(* IEC 61131-3 sources: plc-st-coding-agent/progress/evidence/f14_p1_20261111b/jobs/codex_minimax-m27, 60 files *)

(* ---- public-easy-02.candidate_01.st ---- *)
FUNCTION_BLOCK FB_DualWordEdgeDetection
VAR_INPUT
    value : DWORD;
END_VAR

VAR_OUTPUT
    hasChanged      : BOOL;
    hasRisingEdges  : BOOL;
    risingBits      : DWORD;
    noOfRisingBits  : USINT;
    hasFallingEdges : BOOL;
    fallingBits     : DWORD;
    noOfFallingBits : USINT;
END_VAR

VAR
    prevValue : DWORD;
END_VAR

// Detect if the input value has changed
hasChanged := (value <> prevValue);

// Rising edges: current value bit is 1 AND previous value bit was 0
risingBits := value AND (NOT prevValue);
hasRisingEdges := (risingBits <> 0);

// Falling edges: current value bit is 0 AND previous value bit was 1
fallingBits := (NOT value) AND prevValue;
hasFallingEdges := (fallingBits <> 0);

// Count the number of set bits in risingBits
noOfRisingBits := 0;
IF risingBits.0 THEN noOfRisingBits := noOfRisingBits + 1; END_IF
IF risingBits.1 THEN noOfRisingBits := noOfRisingBits + 1; END_IF
IF risingBits.2 THEN noOfRisingBits := noOfRisingBits + 1; END_IF
IF risingBits.3 THEN noOfRisingBits := noOfRisingBits + 1; END_IF
IF risingBits.4 THEN noOfRisingBits := noOfRisingBits + 1; END_IF
IF risingBits.5 THEN noOfRisingBits := noOfRisingBits + 1; END_IF
IF risingBits.6 THEN noOfRisingBits := noOfRisingBits + 1; END_IF
IF risingBits.7 THEN noOfRisingBits := noOfRisingBits + 1; END_IF
IF risingBits.8 THEN noOfRisingBits := noOfRisingBits + 1; END_IF
IF risingBits.9 THEN noOfRisingBits := noOfRisingBits + 1; END_IF
IF risingBits.10 THEN noOfRisingBits := noOfRisingBits + 1; END_IF
IF risingBits.11 THEN noOfRisingBits := noOfRisingBits + 1; END_IF
IF risingBits.12 THEN noOfRisingBits := noOfRisingBits + 1; END_IF
IF risingBits.13 THEN noOfRisingBits := noOfRisingBits + 1; END_IF
IF risingBits.14 THEN noOfRisingBits := noOfRisingBits + 1; END_IF
IF risingBits.15 THEN noOfRisingBits := noOfRisingBits + 1; END_IF
IF risingBits.16 THEN noOfRisingBits := noOfRisingBits + 1; END_IF
IF risingBits.17 THEN noOfRisingBits := noOfRisingBits + 1; END_IF
IF risingBits.18 THEN noOfRisingBits := noOfRisingBits + 1; END_IF
IF risingBits.19 THEN noOfRisingBits := noOfRisingBits + 1; END_IF
IF risingBits.20 THEN noOfRisingBits := noOfRisingBits + 1; END_IF
IF risingBits.21 THEN noOfRisingBits := noOfRisingBits + 1; END_IF
IF risingBits.22 THEN noOfRisingBits := noOfRisingBits + 1; END_IF
IF risingBits.23 THEN noOfRisingBits := noOfRisingBits + 1; END_IF
IF risingBits.24 THEN noOfRisingBits := noOfRisingBits + 1; END_IF
IF risingBits.25 THEN noOfRisingBits := noOfRisingBits + 1; END_IF
IF risingBits.26 THEN noOfRisingBits := noOfRisingBits + 1; END_IF
IF risingBits.27 THEN noOfRisingBits := noOfRisingBits + 1; END_IF
IF risingBits.28 THEN noOfRisingBits := noOfRisingBits + 1; END_IF
IF risingBits.29 THEN noOfRisingBits := noOfRisingBits + 1; END_IF
IF risingBits.30 THEN noOfRisingBits := noOfRisingBits + 1; END_IF
IF risingBits.31 THEN noOfRisingBits := noOfRisingBits + 1; END_IF

// Count the number of set bits in fallingBits
noOfFallingBits := 0;
IF fallingBits.0 THEN noOfFallingBits := noOfFallingBits + 1; END_IF
IF fallingBits.1 THEN noOfFallingBits := noOfFallingBits + 1; END_IF
IF fallingBits.2 THEN noOfFallingBits := noOfFallingBits + 1; END_IF
IF fallingBits.3 THEN noOfFallingBits := noOfFallingBits + 1; END_IF
IF fallingBits.4 THEN noOfFallingBits := noOfFallingBits + 1; END_IF
IF fallingBits.5 THEN noOfFallingBits := noOfFallingBits + 1; END_IF
IF fallingBits.6 THEN noOfFallingBits := noOfFallingBits + 1; END_IF
IF fallingBits.7 THEN noOfFallingBits := noOfFallingBits + 1; END_IF
IF fallingBits.8 THEN noOfFallingBits := noOfFallingBits + 1; END_IF
IF fallingBits.9 THEN noOfFallingBits := noOfFallingBits + 1; END_IF
IF fallingBits.10 THEN noOfFallingBits := noOfFallingBits + 1; END_IF
IF fallingBits.11 THEN noOfFallingBits := noOfFallingBits + 1; END_IF
IF fallingBits.12 THEN noOfFallingBits := noOfFallingBits + 1; END_IF
IF fallingBits.13 THEN noOfFallingBits := noOfFallingBits + 1; END_IF
IF fallingBits.14 THEN noOfFallingBits := noOfFallingBits + 1; END_IF
IF fallingBits.15 THEN noOfFallingBits := noOfFallingBits + 1; END_IF
IF fallingBits.16 THEN noOfFallingBits := noOfFallingBits + 1; END_IF
IF fallingBits.17 THEN noOfFallingBits := noOfFallingBits + 1; END_IF
IF fallingBits.18 THEN noOfFallingBits := noOfFallingBits + 1; END_IF
IF fallingBits.19 THEN noOfFallingBits := noOfFallingBits + 1; END_IF
IF fallingBits.20 THEN noOfFallingBits := noOfFallingBits + 1; END_IF
IF fallingBits.21 THEN noOfFallingBits := noOfFallingBits + 1; END_IF
IF fallingBits.22 THEN noOfFallingBits := noOfFallingBits + 1; END_IF
IF fallingBits.23 THEN noOfFallingBits := noOfFallingBits + 1; END_IF
IF fallingBits.24 THEN noOfFallingBits := noOfFallingBits + 1; END_IF
IF fallingBits.25 THEN noOfFallingBits := noOfFallingBits + 1; END_IF
IF fallingBits.26 THEN noOfFallingBits := noOfFallingBits + 1; END_IF
IF fallingBits.27 THEN noOfFallingBits := noOfFallingBits + 1; END_IF
IF fallingBits.28 THEN noOfFallingBits := noOfFallingBits + 1; END_IF
IF fallingBits.29 THEN noOfFallingBits := noOfFallingBits + 1; END_IF
IF fallingBits.30 THEN noOfFallingBits := noOfFallingBits + 1; END_IF
IF fallingBits.31 THEN noOfFallingBits := noOfFallingBits + 1; END_IF

// Store current value for next cycle
prevValue := value;

END_FUNCTION_BLOCK

(* ---- public-easy-02.candidate_02.st ---- *)
FUNCTION_BLOCK FB_DualWordEdgeDetection
VAR_INPUT
    value : DWORD;
END_VAR

VAR_OUTPUT
    hasChanged      : BOOL;
    hasRisingEdges  : BOOL;
    risingBits      : DWORD;
    noOfRisingBits  : USINT;
    hasFallingEdges : BOOL;
    fallingBits     : DWORD;
    noOfFallingBits : USINT;
END_VAR

VAR
    prevValue : DWORD;
END_VAR

// Detect if the input value has changed
hasChanged := (value <> prevValue);

// Rising edges: current value bit is 1 AND previous value bit was 0
risingBits := value AND (NOT prevValue);
hasRisingEdges := (risingBits <> 0);

// Falling edges: current value bit is 0 AND previous value bit was 1
fallingBits := (NOT value) AND prevValue;
hasFallingEdges := (fallingBits <> 0);

// Count the number of set bits in risingBits using bit manipulation
noOfRisingBits := 0;
VAR tempRising : DWORD; END_VAR
tempRising := risingBits;
WHILE tempRising <> 0 DO
    noOfRisingBits := noOfRisingBits + 1;
    tempRising := tempRising AND (tempRising - 1); // Clear lowest set bit
END_WHILE

// Count the number of set bits in fallingBits using bit manipulation
noOfFallingBits := 0;
VAR tempFalling : DWORD; END_VAR
tempFalling := fallingBits;
WHILE tempFalling <> 0 DO
    noOfFallingBits := noOfFallingBits + 1;
    tempFalling := tempFalling AND (tempFalling - 1); // Clear lowest set bit
END_WHILE

// Store current value for next cycle
prevValue := value;

END_FUNCTION_BLOCK

(* ---- public-easy-03.candidate_01.st ---- *)
FUNCTION_BLOCK AlarmHandler
VAR_INPUT
    Value       : REAL;
    hiLevel     : REAL;
    loLevel     : REAL;
    hystWindow  : REAL;
END_VAR

VAR_OUTPUT
    hiAlarm     : BOOL;
    loAlarm     : BOOL;
    error       : BOOL;
    status      : WORD;
END_VAR

// Error checking
IF loLevel >= hiLevel THEN
    error := TRUE;
    status := 16#8001;
    RETURN;
END_IF

IF hystWindow >= (hiLevel - loLevel) THEN
    error := TRUE;
    status := 16#8002;
    RETURN;
END_IF

// No error
error := FALSE;
status := 16#0000;

// High alarm with hysteresis
// Trigger: Value > hiLevel
// Reset:   Value < hiLevel - hystWindow
IF Value > hiLevel THEN
    hiAlarm := TRUE;
ELSIF Value < (hiLevel - hystWindow) THEN
    hiAlarm := FALSE;
END_IF

// Low alarm with hysteresis
// Trigger: Value < loLevel
// Reset:   Value > loLevel + hystWindow
IF Value < loLevel THEN
    loAlarm := TRUE;
ELSIF Value > (loLevel + hystWindow) THEN
    loAlarm := FALSE;
END_IF

END_FUNCTION_BLOCK

(* ---- public-easy-03.candidate_02.st ---- *)
FUNCTION_BLOCK AlarmHandler
VAR_INPUT
    Value       : REAL;
    hiLevel     : REAL;
    loLevel     : REAL;
    hystWindow  : REAL;
END_VAR

VAR_OUTPUT
    hiAlarm     : BOOL;
    loAlarm     : BOOL;
    error       : BOOL;
    status      : WORD;
END_VAR

// Error checking
IF loLevel >= hiLevel THEN
    error := TRUE;
    status := 16#8001;
    RETURN;
END_IF

IF hystWindow >= (hiLevel - loLevel) THEN
    error := TRUE;
    status := 16#8002;
    RETURN;
END_IF

// No error - reset all outputs to defined state
error := FALSE;
status := 16#0000;
hiAlarm := FALSE;
loAlarm := FALSE;

// High alarm with hysteresis
// Trigger: Value > hiLevel
// Reset:   Value < hiLevel - hystWindow
IF Value > hiLevel THEN
    hiAlarm := TRUE;
END_IF

// Low alarm with hysteresis
// Trigger: Value < loLevel
// Reset:   Value > loLevel + hystWindow
IF Value < loLevel THEN
    loAlarm := TRUE;
END_IF

END_FUNCTION_BLOCK

(* ---- public-easy-05.candidate_01.st ---- *)
FUNCTION_BLOCK WeldGapAlarm
VAR_INPUT
    Gap_Exceeded    : BOOL;      // Scanner indication that the gap exceeds 1.5 mm
    Weld_E_Stop_NC  : BOOL;      // TRUE = inactive, FALSE = active (emergency stop)
    DebounceTime    : TIME;      // Gap-signal debounce duration during normal monitoring
END_VAR

VAR_OUTPUT
    Operator_Alert         : BOOL;  // Audible and visual alarm command
    Weld_Soft_Start_Active : BOOL;  // Monitoring-inhibition status during 5-second power-up initialization
END_VAR

VAR
    InitTimer    : TON;          // 5-second initialization inhibition timer
    DebounceTmr  : TON;          // Gap signal debounce timer during normal monitoring
    bInitDone    : BOOL;         // Power-up initialization completion flag
END_VAR

    // E-Stop takes highest priority over initialization and normal monitoring
    IF NOT Weld_E_Stop_NC THEN
        Operator_Alert         := FALSE;
        Weld_Soft_Start_Active := FALSE;
        DebounceTmr(IN := FALSE);
        InitTimer(IN := FALSE);
        bInitDone := FALSE;
        RETURN;
    END_IF

    // 5-second initialization inhibition period
    IF NOT bInitDone THEN
        Weld_Soft_Start_Active := TRUE;
        Operator_Alert         := FALSE;
        InitTimer(IN := TRUE, PT := T#5S);

        IF InitTimer.Q THEN
            bInitDone := TRUE;
            InitTimer(IN := FALSE);
        END_IF;

        // During initialization, debounce time does NOT accumulate
        RETURN;
    END_IF;

    // Normal gap monitoring after initialization
    Weld_Soft_Start_Active := FALSE;

    // Debounce logic: alarm only after Gap_Exceeded remains TRUE for DebounceTime
    IF Gap_Exceeded THEN
        DebounceTmr(IN := TRUE, PT := DebounceTime);
        Operator_Alert := DebounceTmr.Q;
    ELSE
        DebounceTmr(IN := FALSE);
        Operator_Alert := FALSE;
    END_IF;

END_FUNCTION_BLOCK

(* ---- public-easy-05.candidate_02.st ---- *)
FUNCTION_BLOCK WeldGapAlarm
VAR_INPUT
    Gap_Exceeded    : BOOL;      // Scanner indication that the gap exceeds 1.5 mm
    Weld_E_Stop_NC  : BOOL;      // TRUE = inactive, FALSE = active (emergency stop)
    DebounceTime    : TIME;      // Gap-signal debounce duration during normal monitoring
END_VAR

VAR_OUTPUT
    Operator_Alert         : BOOL;  // Audible and visual alarm command
    Weld_Soft_Start_Active : BOOL;  // Monitoring-inhibition status during 5-second power-up initialization
END_VAR

VAR
    InitTimer    : TON;          // 5-second initialization inhibition timer
    DebounceTmr  : TON;          // Gap signal debounce timer during normal monitoring
    bInitDone    : BOOL;         // Power-up initialization completion flag
END_VAR

    // E-Stop takes highest priority over initialization and normal monitoring
    IF NOT Weld_E_Stop_NC THEN
        Operator_Alert         := FALSE;
        Weld_Soft_Start_Active := FALSE;
        DebounceTmr(IN := FALSE, R := TRUE);
        InitTimer(IN := FALSE, R := TRUE);
        bInitDone := FALSE;
        RETURN;
    END_IF

    // 5-second initialization inhibition period
    IF NOT bInitDone THEN
        Weld_Soft_Start_Active := TRUE;
        Operator_Alert         := FALSE;
        InitTimer(IN := TRUE, PT := T#5S);

        IF InitTimer.Q THEN
            bInitDone := TRUE;
            InitTimer(IN := FALSE);
        END_IF;

        // During initialization, debounce time does NOT accumulate
        RETURN;
    END_IF;

    // Normal gap monitoring after initialization
    Weld_Soft_Start_Active := FALSE;

    // Debounce logic: alarm only after Gap_Exceeded remains TRUE for DebounceTime
    IF Gap_Exceeded THEN
        DebounceTmr(IN := TRUE, PT := DebounceTime);
        Operator_Alert := DebounceTmr.Q;
    ELSE
        DebounceTmr(IN := FALSE, PT := DebounceTime);  // Reset timer to clear accumulated time
        Operator_Alert := FALSE;
    END_IF;

END_FUNCTION_BLOCK

(* ---- public-easy-06.candidate_02.st ---- *)
FUNCTION_BLOCK AerationBlower
VAR_INPUT
    do_low               : BOOL;
    aeration_e_stop_nc   : BOOL;
END_VAR

VAR_OUTPUT
    blower_run                   : BOOL;
    aeration_blower_cycle_count  : UINT;
END_VAR

VAR
    start_timer        : TON;
    blower_was_running : BOOL;
END_VAR

// Start delay: timer runs while both conditions are met
start_timer(
    IN := do_low AND aeration_e_stop_nc,
    PT := T#5S
);

// Blower runs only when timer elapsed AND conditions remain satisfied
blower_run := start_timer.Q AND do_low AND aeration_e_stop_nc;

// Count FALSE-to-TRUE transitions of blower_run (rising edge)
IF blower_run AND NOT blower_was_running THEN
    aeration_blower_cycle_count := aeration_blower_cycle_count + 1;
END_IF;

// Update edge-detection state for next scan
blower_was_running := blower_run;

END_FUNCTION_BLOCK

(* ---- public-hard-01.candidate_02.st ---- *)
// Material Proportioning Process Control - ST Implementation
FUNCTION_BLOCK MaterialProportioning
VAR_INPUT
    estop            : BOOL;   // Emergency Stop Signal (FALSE = triggered)
    opeMode          : BOOL;   // Operation Mode (FALSE = Manual, TRUE = Auto)
    valveAStart      : BOOL;   // Valve A Start Button
    valveBStart      : BOOL;   // Valve B Start Button
    valveCStart      : BOOL;   // Valve C Start Button
    valveDStart      : BOOL;   // Valve D Start Button
    mixMotorStart    : BOOL;   // Mixing Motor Start Button
    autoStart        : BOOL;   // Automatic Start Button
    processMode      : BOOL;   // Process Mode (FALSE = Basic, TRUE = Extended)
    levelSensor      : INT;    // Liquid Level Sensor (unit: cm)
    mixMotorComplete : BOOL;   // Mixing Complete Signal
END_VAR

VAR_OUTPUT
    valveARun  : BOOL;   // Valve A Run Command
    valveBRun  : BOOL;   // Valve B Run Command
    valveCRun  : BOOL;   // Valve C Run Command
    valveDRun  : BOOL;   // Valve D Run Command
    mixMotorRun: BOOL;   // Mixing Motor Run Command
END_VAR

VAR
    prevValveAStart   : BOOL;   // Previous state for edge detection
    prevValveBStart   : BOOL;
    prevValveCStart   : BOOL;
    prevValveDStart   : BOOL;
    prevMixMotorStart : BOOL;
    prevAutoStart     : BOOL;
    autoState : INT;     // 0=IDLE, 1=FILL_A, 2=FILL_B, 3=MIX_BASIC,
                         // 4=FILL_C, 5=MIX_EXT, 6=DRAIN
END_VAR

VAR CONSTANT
    STATE_IDLE      : INT := 0;
    STATE_FILL_A    : INT := 1;
    STATE_FILL_B    : INT := 2;
    STATE_MIX_BASIC : INT := 3;
    STATE_FILL_C    : INT := 4;
    STATE_MIX_EXT   : INT := 5;
    STATE_DRAIN     : INT := 6;
END_VAR

// ============================================================================
// Main Control Logic
// ============================================================================

// ---------------------------------------------------------------------------
// Emergency Stop Logic
// When estop=FALSE, all equipment stops immediately
// ---------------------------------------------------------------------------
IF NOT estop THEN
    valveARun  := FALSE;
    valveBRun  := FALSE;
    valveCRun  := FALSE;
    valveDRun  := FALSE;
    mixMotorRun:= FALSE;
    autoState  := STATE_IDLE;

    prevValveAStart   := FALSE;
    prevValveBStart   := FALSE;
    prevValveCStart   := FALSE;
    prevValveDStart   := FALSE;
    prevMixMotorStart := FALSE;
    prevAutoStart     := FALSE;
    RETURN;
END_IF

// ---------------------------------------------------------------------------
// Mode Selection: Manual vs Automatic
// ---------------------------------------------------------------------------
IF NOT opeMode THEN
    // MANUAL OPERATION MODE
    // Toggle each device on rising edge of corresponding button

    IF valveAStart AND NOT prevValveAStart THEN
        valveARun := NOT valveARun;
    END_IF;
    prevValveAStart := valveAStart;

    IF valveBStart AND NOT prevValveBStart THEN
        valveBRun := NOT valveBRun;
    END_IF;
    prevValveBStart := valveBStart;

    IF valveCStart AND NOT prevValveCStart THEN
        valveCRun := NOT valveCRun;
    END_IF;
    prevValveCStart := valveCStart;

    IF valveDStart AND NOT prevValveDStart THEN
        valveDRun := NOT valveDRun;
    END_IF;
    prevValveDStart := valveDStart;

    IF mixMotorStart AND NOT prevMixMotorStart THEN
        mixMotorRun := NOT mixMotorRun;
    END_IF;
    prevMixMotorStart := mixMotorStart;

ELSE
    // AUTOMATIC OPERATION MODE

    valveARun  := FALSE;
    valveBRun  := FALSE;
    valveCRun  := FALSE;
    valveDRun  := FALSE;
    mixMotorRun:= FALSE;

    IF autoStart AND NOT prevAutoStart THEN
        IF autoState = STATE_IDLE THEN
            autoState := STATE_FILL_A;
        END_IF;
    END_IF;
    prevAutoStart := autoStart;

    CASE autoState OF

        STATE_IDLE:
            valveARun  := FALSE;
            valveBRun  := FALSE;
            valveCRun  := FALSE;
            valveDRun  := FALSE;
            mixMotorRun:= FALSE;

        STATE_FILL_A:
            valveARun := TRUE;
            IF levelSensor >= 50 THEN
                valveARun := FALSE;
                autoState := STATE_FILL_B;
            END_IF;

        STATE_FILL_B:
            valveBRun := TRUE;
            IF levelSensor >= 80 THEN
                valveBRun := FALSE;
                IF NOT processMode THEN
                    autoState := STATE_MIX_BASIC;
                ELSE
                    autoState := STATE_FILL_C;
                END_IF;
            END_IF;

        STATE_MIX_BASIC:
            mixMotorRun := TRUE;
            IF mixMotorComplete THEN
                mixMotorRun := FALSE;
                autoState := STATE_DRAIN;
            END_IF;

        STATE_FILL_C:
            valveCRun := TRUE;
            IF levelSensor >= 100 THEN
                valveCRun := FALSE;
                autoState := STATE_MIX_EXT;
            END_IF;

        STATE_MIX_EXT:
            mixMotorRun := TRUE;
            IF mixMotorComplete THEN
                mixMotorRun := FALSE;
                autoState := STATE_DRAIN;
            END_IF;

        STATE_DRAIN:
            valveDRun := TRUE;
            IF levelSensor < 10 THEN
                valveDRun := FALSE;
                autoState := STATE_IDLE;
            END_IF;

    END_CASE;

END_IF;

END_FUNCTION_BLOCK

PROGRAM PLC_PRG
VAR
    inst : MaterialProportioning;
END_VAR

inst(
    estop            := estop,
    opeMode          := opeMode,
    valveAStart      := valveAStart,
    valveBStart      := valveBStart,
    valveCStart      := valveCStart,
    valveDStart      := valveDStart,
    mixMotorStart    := mixMotorStart,
    autoStart        := autoStart,
    processMode      := processMode,
    levelSensor      := levelSensor,
    mixMotorComplete := mixMotorComplete,
    valveARun        => valveARun,
    valveBRun        => valveBRun,
    valveCRun        => valveCRun,
    valveDRun        => valveDRun,
    mixMotorRun      => mixMotorRun
);
END_PROGRAM

(* ---- public-hard-04.candidate_02.st ---- *)
FUNCTION_BLOCK FB_FIFO
VAR_INPUT
    enqueue : BOOL;
    dequeue : BOOL;
    reset   : BOOL;
END_VAR

VAR_OUTPUT
    elementCount : DINT;
    status       : WORD;
END_VAR

VAR_IN_OUT
    item   : VARIANT;
    buffer : VARIANT;
END_VAR

VAR
    _head         : DINT := 0;
    _tail         : DINT := 0;
    _elementCount : DINT := 0;
    _capacity     : DINT;
    _elementSize  : DINT;
    _prevEnqueue  : BOOL := FALSE;
    _prevDequeue  : BOOL := FALSE;
    _initialized  : BOOL := FALSE;
END_VAR

// Initialization
IF NOT _initialized THEN
    VAR
        bufType : REF_TO ANY;
        capacity : DINT;
    END_VAR

    bufType REF= buffer;

    IF __ISVALIDREF(bufType) THEN
        capacity := bufType.GetUpperBound(1) + 1;
        _capacity := capacity;
        _elementSize := bufType.GetSize() / _capacity;
        _initialized := TRUE;
    END_IF;

    elementCount := 0;
    status := 16#0000;
    RETURN;
END_IF;

// Reset handling (highest priority)
IF reset THEN
    _head := 0;
    _tail := 0;
    _elementCount := 0;
    elementCount := 0;
    status := 16#0000;
    _prevEnqueue := FALSE;
    _prevDequeue := FALSE;
    RETURN;
END_IF;

// Rising edge detection
VAR
    enqueueRising : BOOL;
    dequeueRising : BOOL;
END_VAR

enqueueRising := enqueue AND NOT _prevEnqueue;
dequeueRising := dequeue AND NOT _prevDequeue;

_prevEnqueue := enqueue;
_prevDequeue := dequeue;

// Dequeue request (rising edge, queue not empty)
IF dequeueRising AND _elementCount > 0 THEN
    VAR
        pSrc     : POINTER TO BYTE;
        pDest    : POINTER TO BYTE;
        srcAdr   : LWORD;
        destAdr  : LWORD;
        zeroBuf  : ARRAY[0..255] OF BYTE;
    END_VAR

    srcAdr := __GET_VAR_DATA_REF(buffer).ADR + (_head * _elementSize);
    destAdr := __GET_VAR_DATA_REF(item).ADR;

    MemMove(TO_PTR(srcAdr), TO_PTR(destAdr), _elementSize);

    MemSet(zeroBuf, 0, SIZEOF(zeroBuf));
    MemMove(zeroBuf, TO_PTR(srcAdr), _elementSize);

    _head := (_head + 1) MOD _capacity;
    _elementCount := _elementCount - 1;
    elementCount := _elementCount;
    status := 16#0000;

// Enqueue request (rising edge, queue not full)
ELSIF enqueueRising AND _elementCount < _capacity THEN
    VAR
        pDest   : POINTER TO BYTE;
        pSrc    : POINTER TO BYTE;
        destAdr : LWORD;
        srcAdr  : LWORD;
    END_VAR

    destAdr := __GET_VAR_DATA_REF(buffer).ADR + (_tail * _elementSize);
    srcAdr := __GET_VAR_DATA_REF(item).ADR;

    MemMove(TO_PTR(srcAdr), TO_PTR(destAdr), _elementSize);

    _tail := (_tail + 1) MOD _capacity;
    _elementCount := _elementCount + 1;
    elementCount := _elementCount;
    status := 16#0000;

// Dequeue rejected: empty queue
ELSIF dequeueRising AND _elementCount = 0 THEN
    status := 16#8001;

// Enqueue rejected: full queue
ELSIF enqueueRising AND _elementCount >= _capacity THEN
    status := 16#8002;

// Idle (no rising edge or other condition)
ELSE
    status := 16#0000;
END_IF;
END_FUNCTION_BLOCK

(* ---- public-medium-01.candidate_02.st ---- *)
FUNCTION_BLOCK FB_MultiPumpControl
VAR_INPUT
    mode    : BOOL;  // FALSE: Manual mode, TRUE: Automatic mode
    start   : BOOL;  // Start button
    stop    : BOOL;  // Stop button
END_VAR

VAR_IN_OUT
    pumpGroup   : ARRAY[1..5] OF ST_Pump;
END_VAR

VAR
    startOld    : BOOL := FALSE;
    stopOld     : BOOL := FALSE;
    startEdge   : BOOL;
    stopEdge    : BOOL;
    i           : INT;
    runCount    : INT;
    tempPump    : ST_Pump;
    sorted      : BOOL := FALSE;
    priorities  : ARRAY[1..5] OF INT;
END_VAR

// Detect rising edges
startEdge := start AND NOT startOld;
stopEdge  := stop  AND NOT stopOld;
startOld  := start;
stopOld   := stop;

// Stop all pumps when stop is pressed
IF stopEdge THEN
    FOR i := 1 TO 5 DO
        pumpGroup[i].RunComd := FALSE;
    END_FOR
    sorted := FALSE;
    RETURN;
END_IF

// Start pumps when start is pressed
IF startEdge THEN
    IF mode = FALSE THEN
        // Manual mode: start pumps based on selection
        FOR i := 1 TO 5 DO
            IF pumpGroup[i].selection THEN
                pumpGroup[i].RunComd := TRUE;
            END_IF
        END_FOR
    ELSE
        // Automatic mode: select top 3 by priority (bubble sort)
        // Store priorities
        FOR i := 1 TO 5 DO
            priorities[i] := pumpGroup[i].priority;
        END_FOR

        // Bubble sort priorities and rearrange pumpGroup accordingly
        FOR i := 1 TO 5 DO
            tempPump := pumpGroup[i];
        END_FOR

        // Sort by priority descending
        FOR i := 1 TO 4 DO
            IF priorities[i] < priorities[i+1] THEN
                // Swap priorities
                tempPump := pumpGroup[i];
                pumpGroup[i] := pumpGroup[i+1];
                pumpGroup[i+1] := tempPump;

                // Update priority array
                priorities[i] := pumpGroup[i].priority;
                priorities[i+1] := pumpGroup[i+1].priority;
            END_IF
        END_FOR

        // Select top 3 pumps
        runCount := 0;
        FOR i := 1 TO 5 DO
            IF runCount < 3 THEN
                pumpGroup[i].RunComd := TRUE;
                runCount := runCount + 1;
            ELSE
                pumpGroup[i].RunComd := FALSE;
            END_IF
        END_FOR

        sorted := TRUE;
    END_IF
END_IF
END_FUNCTION_BLOCK

(* ---- public-medium-02.candidate_01.st ---- *)
FUNCTION_BLOCK FB_AnalogBatchProcess
VAR_INPUT
    count : DINT;
END_VAR

VAR_IN_OUT
    analogValues : ARRAY[*] OF INT;
    channels     : ARRAY[*] OF ST_AnalogChannel;
END_VAR

VAR
    i           : DINT;
    idx         : DINT;
    rawValue    : INT;
    channel     : REF_TO ST_AnalogChannel;
END_VAR

// Process each channel by ordinal position
FOR i := 0 TO count - 1 DO
    idx := LOWER_BOUND(channels, 1) + i;
    channel := REF(channels[idx]);

    // Skip disabled channels
    IF NOT channel.enable THEN
        CONTINUE;
    END_IF

    // Default success status
    channel.retVal := 16#0000;

    // Validate hiLIM > loLIM
    IF channel.hiLIM <= channel.loLIM THEN
        channel.retVal := 16#8002;
        CONTINUE;
    END_IF

    // Get raw analog value (read-only)
    rawValue := analogValues[LOWER_BOUND(analogValues, 1) + i];

    // Perform conversion based on measuringMode
    CASE channel.measuringMode OF
        0: // Non-temperature linear scaling
            IF channel.bipolar THEN
                // Bipolar: map -27648..27648 to loLIM..hiLIM
                channel.outputValue := (INT_TO_REAL(rawValue) + 27648.0) / 55296.0 * (channel.hiLIM - channel.loLIM) + channel.loLIM;
            ELSE
                // Unipolar: map 0..27648 to loLIM..hiLIM
                channel.outputValue := INT_TO_REAL(rawValue) / 27648.0 * (channel.hiLIM - channel.loLIM) + channel.loLIM;
            END_IF;

        1: // Standard temperature: outputValue = raw / 10
            channel.outputValue := INT_TO_REAL(rawValue) / 10.0;

        2: // Climatic temperature: outputValue = raw / 100
            channel.outputValue := INT_TO_REAL(rawValue) / 100.0;

    ELSE
        // Invalid measuringMode
        channel.retVal := 16#8001;
    END_CASE;
END_FOR;

END_FUNCTION_BLOCK

(* ---- public-medium-02.candidate_02.st ---- *)
FUNCTION_BLOCK FB_AnalogBatchProcess
VAR_INPUT
    count : DINT;
END_VAR

VAR_IN_OUT
    analogValues : ARRAY[*] OF INT;
    channels     : ARRAY[*] OF ST_AnalogChannel;
END_VAR

VAR
    i           : DINT;
    idx         : DINT;
    rawValue    : INT;
    validInput  : BOOL;
END_VAR

i := 0;
WHILE i < count DO
    idx := LOWER_BOUND(channels, 1) + i;

    // Check if channel is enabled
    IF channels[idx].enable THEN
        // Default success status
        channels[idx].retVal := 16#0000;

        // Validate hiLIM > loLIM
        IF channels[idx].hiLIM > channels[idx].loLIM THEN
            // Get raw analog value
            rawValue := analogValues[LOWER_BOUND(analogValues, 1) + i];

            // Perform conversion based on measuringMode
            CASE channels[idx].measuringMode OF
                0: // Non-temperature linear scaling
                    IF channels[idx].bipolar THEN
                        // Bipolar: map -27648..27648 to loLIM..hiLIM
                        channels[idx].outputValue := (INT_TO_REAL(rawValue) + 27648.0) / 55296.0 * (channels[idx].hiLIM - channels[idx].loLIM) + channels[idx].loLIM;
                    ELSE
                        // Unipolar: map 0..27648 to loLIM..hiLIM
                        channels[idx].outputValue := INT_TO_REAL(rawValue) / 27648.0 * (channels[idx].hiLIM - channels[idx].loLIM) + channels[idx].loLIM;
                    END_IF;

                1: // Standard temperature: outputValue = raw / 10
                    channels[idx].outputValue := INT_TO_REAL(rawValue) / 10.0;

                2: // Climatic temperature: outputValue = raw / 100
                    channels[idx].outputValue := INT_TO_REAL(rawValue) / 100.0;

            ELSE
                // Invalid measuringMode
                channels[idx].retVal := 16#8001;
            END_CASE;
        ELSE
            // hiLIM <= loLIM error
            channels[idx].retVal := 16#8002;
        END_IF;
    END_IF;

    i := i + 1;
END_WHILE;

END_FUNCTION_BLOCK

(* ---- public-medium-04.candidate_01.st ---- *)
FUNCTION_BLOCK FB_TemperatureControl
VAR_INPUT
    TemperatureSensorInput : REAL;
    SetTemperature         : REAL;
END_VAR

VAR_OUTPUT
    CurrentTemperature : REAL;
    SetTempDisplay     : REAL;
    HeaterStatus       : BOOL;
    OverheatProtection : BOOL;
    HeaterOutput       : BOOL;
END_VAR

VAR
    // Internal variables
    rCurrentTemperature  : REAL := 0.0;
    rSetTemperature      : REAL := 0.0;
    bHeaterOn            : BOOL := FALSE;
    bOverheatProtection  : BOOL := FALSE;
    bSensorFault         : BOOL := FALSE;

    // Timer for heater on-time monitoring
    HeaterOnTimer        : TON;
    // Timer for overheat protection cooldown
    OverheatCooldownTimer: TON;

    // Constants
    MAX_HEATER_ON_TIME   : TIME := T#5S;
    OVERHEAT_COOLDOWN    : TIME := T#3S;
    MIN_SENSOR_VALUE     : REAL := 0.0;
    MAX_SENSOR_VALUE     : REAL := 100.0;
END_VAR

//============================================================================
// Temperature Logic Control - Main Program
//============================================================================

// Update internal temperature values from inputs
rCurrentTemperature := TemperatureSensorInput;
rSetTemperature     := SetTemperature;

// Update output displays
CurrentTemperature := rCurrentTemperature;
SetTempDisplay     := rSetTemperature;
HeaterStatus       := bHeaterOn;
OverheatProtection := bOverheatProtection;

//============================================================================
// Sensor Fault Detection
// If temperature is outside valid range (0-100), trigger sensor fault
//============================================================================
bSensorFault := (rCurrentTemperature < MIN_SENSOR_VALUE) OR
                (rCurrentTemperature > MAX_SENSOR_VALUE);

IF bSensorFault THEN
    // Sensor fault: turn off heater immediately
    bHeaterOn          := FALSE;
    HeaterOutput       := FALSE;
    bOverheatProtection := TRUE;

    // Reset heater on timer when heater is off
    HeaterOnTimer(IN := FALSE);

    // Return early - no temperature control during sensor fault
    RETURN;
END_IF;

//============================================================================
// Overheat Protection Check
// If protection is active, must wait for cooldown period before reset
//============================================================================
IF bOverheatProtection THEN
    // Start or continue cooldown timer
    OverheatCooldownTimer(IN := TRUE, PT := OVERHEAT_COOLDOWN);

    // Check if cooldown period has elapsed
    IF OverheatCooldownTimer.Q THEN
        // Cooldown complete - reset overheat protection
        bOverheatProtection        := FALSE;
        OverheatCooldownTimer(IN := FALSE);
    END_IF;

    // Keep heater off during overheat protection
    bHeaterOn := FALSE;
    HeaterOutput := FALSE;

    // Return early - no temperature control during overheat protection
    RETURN;
ELSE
    // Reset cooldown timer when protection is not active
    OverheatCooldownTimer(IN := FALSE);
END_IF;

//============================================================================
// Temperature Control Logic
// Compare actual temperature with set temperature
//============================================================================
IF rCurrentTemperature < rSetTemperature THEN
    // Temperature below setpoint - turn ON heater
    bHeaterOn := TRUE;
ELSIF rCurrentTemperature >= rSetTemperature THEN
    // Temperature at or above setpoint - turn OFF heater
    bHeaterOn := FALSE;
END_IF;

//============================================================================
// Heater Output Control
//============================================================================
HeaterOutput := bHeaterOn;

//============================================================================
// Heater On-Time Monitoring for Overheat Protection
// If heater runs continuously for more than 5 seconds, trigger protection
//============================================================================
IF bHeaterOn THEN
    // Start or continue the heater on-time timer
    HeaterOnTimer(IN := TRUE, PT := MAX_HEATER_ON_TIME);

    // Check if timer has elapsed (heater on for too long)
    IF HeaterOnTimer.Q THEN
        // Overheat protection triggered
        bHeaterOn           := FALSE;
        bOverheatProtection := TRUE;
        HeaterOutput        := FALSE;

        // Reset heater on timer
        HeaterOnTimer(IN := FALSE);
    END_IF;
ELSE
    // Heater is off - reset the timer
    HeaterOnTimer(IN := FALSE);
END_IF;

END_FUNCTION_BLOCK

(* ---- public-medium-04.candidate_02.st ---- *)
FUNCTION_BLOCK FB_TemperatureControl
VAR_INPUT
    TemperatureSensorInput : REAL;
    SetTemperature         : REAL;
END_VAR

VAR_OUTPUT
    CurrentTemperature : REAL;
    SetTempDisplay     : REAL;
    HeaterStatus       : BOOL;
    OverheatProtection : BOOL;
    HeaterOutput       : BOOL;
END_VAR

VAR
    bHeaterOn            : BOOL := FALSE;
    bOverheatProtection  : BOOL := FALSE;

    HeaterOnTimer        : TON;
    OverheatCooldownTimer: TON;

    MAX_HEATER_ON_TIME   : TIME := T#5S;
    OVERHEAT_COOLDOWN    : TIME := T#3S;
END_VAR

//============================================================================
// Main Control Logic
//============================================================================

// Sensor Fault Detection (0-100 valid range)
IF (TemperatureSensorInput < 0.0) OR (TemperatureSensorInput > 100.0) THEN
    // Sensor fault: disable heater and activate protection
    bHeaterOn := FALSE;
    bOverheatProtection := TRUE;
    HeaterOnTimer(IN := FALSE);
END_IF

// Overheat Protection Logic
IF bOverheatProtection THEN
    OverheatCooldownTimer(IN := TRUE, PT := OVERHEAT_COOLDOWN);

    IF OverheatCooldownTimer.Q THEN
        bOverheatProtection := FALSE;
        OverheatCooldownTimer(IN := FALSE);
    END_IF;

    bHeaterOn := FALSE;
ELSE
    OverheatCooldownTimer(IN := FALSE);

    // Temperature Control (only when no protection active)
    IF TemperatureSensorInput < SetTemperature THEN
        bHeaterOn := TRUE;
    ELSE
        bHeaterOn := FALSE;
    END_IF;
END_IF;

// Heater On-Time Monitoring
IF bHeaterOn THEN
    HeaterOnTimer(IN := TRUE, PT := MAX_HEATER_ON_TIME);

    IF HeaterOnTimer.Q THEN
        bHeaterOn := FALSE;
        bOverheatProtection := TRUE;
        HeaterOnTimer(IN := FALSE);
    END_IF;
ELSE
    HeaterOnTimer(IN := FALSE);
END_IF;

//============================================================================
// Update All Outputs (at the end, after all logic)
//============================================================================
CurrentTemperature := TemperatureSensorInput;
SetTempDisplay     := SetTemperature;
HeaterStatus       := bHeaterOn;
OverheatProtection := bOverheatProtection;
HeaterOutput       := bHeaterOn;

END_FUNCTION_BLOCK

(* ---- public-medium-06.candidate_02.st ---- *)
FUNCTION_BLOCK SlabThicknessMonitor
VAR_INPUT
    THICKNESS_FAULT        : BOOL;
    THICKNESS_SIGNAL_VALID : BOOL;
    cutting_run            : BOOL;
    faulttimestamp         : DINT;
    cycletime              : TIME;
END_VAR

VAR_OUTPUT
    THICKNESS_ALARM           : BOOL;
    slab_fault_counter        : UINT;
    slab_runtime_accumulator  : LTIME;
    slab_fault_history        : ARRAY[0..4] OF DINT;
END_VAR

VAR
    AlarmHoldTimer   : TON;
    FaultWasActive   : BOOL;
    PowerUpComplete  : BOOL;
    i                : INT;
END_VAR

IF NOT PowerUpComplete THEN
    THICKNESS_ALARM           := FALSE;
    slab_fault_counter        := 0;
    slab_runtime_accumulator  := LTIME#0s;

    FOR i := 0 TO 4 DO
        slab_fault_history[i] := 0;
    END_FOR

    FaultWasActive  := FALSE;
    PowerUpComplete := TRUE;
END_IF

IF NOT THICKNESS_SIGNAL_VALID THEN
    THICKNESS_ALARM := FALSE;
    AlarmHoldTimer(IN := FALSE);
    FaultWasActive  := FALSE;
ELSE
    AlarmHoldTimer(IN := THICKNESS_FAULT, PT := T#500ms);
    THICKNESS_ALARM := THICKNESS_FAULT OR AlarmHoldTimer.Q;

    IF THICKNESS_FAULT AND NOT FaultWasActive THEN
        slab_fault_counter        := slab_fault_counter + 1;
        slab_fault_history[4]     := slab_fault_history[3];
        slab_fault_history[3]     := slab_fault_history[2];
        slab_fault_history[2]     := slab_fault_history[1];
        slab_fault_history[1]     := slab_fault_history[0];
        slab_fault_history[0]     := faulttimestamp;
    END_IF;

    FaultWasActive := THICKNESS_FAULT;

    IF cutting_run AND NOT THICKNESS_FAULT THEN
        slab_runtime_accumulator := slab_runtime_accumulator + cycletime;
    END_IF
END_IF

END_FUNCTION_BLOCK

(* ---- public-medium-07.candidate_02.st ---- *)
FUNCTION_BLOCK HVAC_Control
VAR_INPUT
    OCCUPANCY_DETECTED    : BOOL;
    ENERGY_SAVING_MODE    : BOOL;
    HVAC_MODE_SELECTOR    : INT;
END_VAR

VAR_OUTPUT
    SUPPLY_FAN_RUN        : BOOL := FALSE;
    TEMP_SETPOINT_ADJUST  : INT := 0;
END_VAR

VAR
    occupancy_delay_timer : TON;
END_VAR

// Fan control with 30-second delay
IF OCCUPANCY_DETECTED AND (HVAC_MODE_SELECTOR <> 3) THEN
    occupancy_delay_timer(IN := TRUE, PT := T#30S);
    IF occupancy_delay_timer.Q THEN
        SUPPLY_FAN_RUN := TRUE;
    ELSE
        SUPPLY_FAN_RUN := FALSE;
    END_IF;
ELSE
    occupancy_delay_timer(IN := FALSE);
    SUPPLY_FAN_RUN := FALSE;
END_IF;

// Temperature setpoint adjustment per mode
CASE HVAC_MODE_SELECTOR OF
    0: // Auto
        IF OCCUPANCY_DETECTED THEN
            TEMP_SETPOINT_ADJUST := 0;
        ELSE
            TEMP_SETPOINT_ADJUST := BOOL_TO_INT(ENERGY_SAVING_MODE) + 2;
        END_IF;
    1: // Comfort
        IF OCCUPANCY_DETECTED THEN
            TEMP_SETPOINT_ADJUST := 0;
        ELSE
            TEMP_SETPOINT_ADJUST := 1;
        END_IF;
    2: // Economy
        IF OCCUPANCY_DETECTED THEN
            TEMP_SETPOINT_ADJUST := 0;
        ELSE
            TEMP_SETPOINT_ADJUST := 4;
        END_IF;
    3: // Night
        TEMP_SETPOINT_ADJUST := 4;
    ELSE
        TEMP_SETPOINT_ADJUST := 0;
END_CASE;

// Clamp to ±4°C
IF TEMP_SETPOINT_ADJUST > 4 THEN
    TEMP_SETPOINT_ADJUST := 4;
ELSIF TEMP_SETPOINT_ADJUST < -4 THEN
    TEMP_SETPOINT_ADJUST := -4;
END_IF;

END_FUNCTION_BLOCK

(* ---- public-medium-08.candidate_01.st ---- *)
FUNCTION_BLOCK FB_IPv4Parse
    VAR_INPUT
        ipText : STRING(254);
    END_VAR
    VAR_OUTPUT
        ipValue : UDINT;
    END_VAR
    VAR
        pos : INT;
        segmentStart : INT;
        segmentLen : INT;
        segmentCount : INT;
        value : INT;
        ch : CHAR;
        textLen : INT;
    END_VAR

    ipValue := 0;
    textLen := LEN(ipText);
    pos := 1;
    segmentCount := 0;

    // Skip leading whitespace
    WHILE (pos <= textLen) AND (MID(ipText, 1, pos) = ' ') DO
        pos := pos + 1;
    END_WHILE;

    // Parse up to 4 segments
    WHILE (segmentCount < 4) AND (pos <= textLen) DO
        segmentStart := pos;
        segmentLen := 0;

        // Collect digits for current segment
        WHILE (pos <= textLen) DO
            ch := MID(ipText, 1, pos);
            IF ch = '.' THEN
                EXIT;
            END_IF;
            IF (ch < '0') OR (ch > '9') THEN
                ipValue := 0;
                RETURN;
            END_IF;
            segmentLen := segmentLen + 1;
            pos := pos + 1;
        END_WHILE;

        // Check segment length (1-3 digits for valid 0-255)
        IF segmentLen < 1 OR segmentLen > 3 THEN
            ipValue := 0;
            RETURN;
        END_IF;

        // Parse segment value
        value := 0;
        FOR pos := segmentStart TO segmentStart + segmentLen - 1 DO
            ch := MID(ipText, 1, pos);
            value := value * 10 + (ch - '0');
        END_FOR;

        // Validate segment range
        IF value > 255 THEN
            ipValue := 0;
            RETURN;
        END_IF;

        // Accumulate result in network byte order
        ipValue := (ipValue << 8) OR TO_UDINT(value);
        segmentCount := segmentCount + 1;

        // Skip the dot separator if present
        IF (pos <= textLen) AND (MID(ipText, 1, pos) = '.') THEN
            pos := pos + 1;
        END_IF;
    END_WHILE;

    // Validate we have exactly 4 segments
    IF segmentCount <> 4 THEN
        ipValue := 0;
        RETURN;
    END_IF;

    // Skip trailing whitespace
    WHILE (pos <= textLen) AND (MID(ipText, 1, pos) = ' ') DO
        pos := pos + 1;
    END_WHILE;

    // If there's more content after the 4 segments (other than whitespace), it's invalid
    IF pos <= textLen THEN
        ipValue := 0;
        RETURN;
    END_IF;

END_FUNCTION_BLOCK

(* ---- public-medium-08.candidate_02.st ---- *)
FUNCTION_BLOCK FB_IPv4Parse
    VAR_INPUT
        ipText : STRING(254);
    END_VAR
    VAR_OUTPUT
        ipValue : UDINT;
    END_VAR
    VAR
        i       : INT;
        pos     : INT;
        start   : INT;
        len     : INT;
        cnt     : INT;
        val     : INT;
        c       : CHAR;
        txtLen  : INT;
        tempPos : INT;
    END_VAR

    ipValue := 0;
    txtLen  := LEN(ipText);
    pos     := 1;
    cnt     := 0;

    // Parse up to 4 segments
    WHILE (cnt < 4) AND (pos <= txtLen) DO
        start := pos;
        len   := 0;

        // Collect digits
        WHILE (pos <= txtLen) DO
            c := MID(ipText, 1, pos);
            IF c = '.' THEN
                EXIT;
            END_IF;
            IF (c < '0') OR (c > '9') THEN
                ipValue := 0;
                RETURN;
            END_IF;
            len := len + 1;
            pos := pos + 1;
        END_WHILE;

        // Check segment length
        IF len < 1 OR len > 3 THEN
            ipValue := 0;
            RETURN;
        END_IF;

        // Parse value
        val := 0;
        tempPos := start;
        FOR i := 1 TO len DO
            c := MID(ipText, 1, tempPos);
            val := val * 10 + (c - '0');
            tempPos := tempPos + 1;
        END_FOR;

        // Range check
        IF val > 255 THEN
            ipValue := 0;
            RETURN;
        END_IF;

        // Accumulate in network byte order (MSB first)
        ipValue := (ipValue * 256) OR TO_UDINT(val);
        cnt := cnt + 1;

        // Skip dot
        IF (pos <= txtLen) AND (MID(ipText, 1, pos) = '.') THEN
            pos := pos + 1;
        END_IF;
    END_WHILE;

    // Must have exactly 4 segments
    IF cnt <> 4 THEN
        ipValue := 0;
        RETURN;
    END_IF;

    // Trailing chars (after dots/skipped) not allowed
    IF pos <= txtLen THEN
        c := MID(ipText, 1, pos);
        IF c <> ' ' AND c <> '' THEN
            ipValue := 0;
            RETURN;
        END_IF;
    END_IF;

END_FUNCTION_BLOCK

(* ---- self-easy-01.candidate_01.st ---- *)
FUNCTION_BLOCK FB
VAR_INPUT
    enable    : BOOL;
    values    : ARRAY[1..8] OF INT;
    count     : INT;
    avgEnable : BOOL;
END_VAR

VAR_OUTPUT
    avgOut : REAL;
END_VAR

VAR
    prev_avgOut : REAL;
END_VAR

IF enable AND avgEnable AND count > 0 THEN
    VAR
        sum : LINT;
        n   : INT;
    END_VAR

    sum := 0;
    IF count > 8 THEN
        n := 8;
    ELSE
        n := count;
    END_IF;

    CASE n OF
        8: sum := sum + values[8];
        7: sum := sum + values[7];
        6: sum := sum + values[6];
        5: sum := sum + values[5];
        4: sum := sum + values[4];
        3: sum := sum + values[3];
        2: sum := sum + values[2];
        1: sum := sum + values[1];
    END_CASE;

    avgOut := LINT_TO_REAL(sum) / INT_TO_REAL(n);
    prev_avgOut := avgOut;
ELSE
    avgOut := prev_avgOut;
END_IF
END_FUNCTION_BLOCK

(* ---- self-easy-01.candidate_02.st ---- *)
FUNCTION_BLOCK FB
VAR_INPUT
    enable    : BOOL;
    values    : ARRAY[1..8] OF INT;
    count     : INT;
    avgEnable : BOOL;
END_VAR

VAR_OUTPUT
    avgOut : REAL;
END_VAR

VAR
    prev_avgOut : REAL;
    sum         : LINT;
    n           : INT;
END_VAR

IF enable AND avgEnable AND count > 0 THEN
    sum := 0;
    IF count > 8 THEN
        n := 8;
    ELSE
        n := count;
    END_IF;

    CASE n OF
        8: sum := sum + values[8];
        7: sum := sum + values[7];
        6: sum := sum + values[6];
        5: sum := sum + values[5];
        4: sum := sum + values[4];
        3: sum := sum + values[3];
        2: sum := sum + values[2];
        1: sum := sum + values[1];
    END_CASE;

    avgOut := LINT_TO_REAL(sum) / INT_TO_REAL(n);
    prev_avgOut := avgOut;
ELSE
    avgOut := prev_avgOut;
END_IF
END_FUNCTION_BLOCK

(* ---- self-easy-02.candidate_01.st ---- *)
FUNCTION_BLOCK FB
VAR_INPUT
    tankLevel    : REAL;      // 储罐液位百分比 0..100
    outletFlow   : REAL;      // 出口流量 m³/h (预留观测接口)
    inletPermit  : BOOL;      // 进料许可
    resetBtn     : BOOL;      // 复位按钮
END_VAR
VAR_OUTPUT
    pumpRun         : BOOL;   // 进料泵运行命令
    alarmHigh       : BOOL;   // 高液位报警
    alarmLow        : BOOL;   // 低液位报警
    outletValveOpen : BOOL;   // 出口阀开命令
END_VAR
VAR
    prevResetBtn : BOOL := FALSE;  // 上拍复位按钮状态
END_VAR

    // 检测复位按钮上升沿：FALSE -> TRUE
    VAR tempRising : BOOL;
    tempRising := resetBtn AND NOT prevResetBtn;

    // --- 高液位报警逻辑 ---
    // 危险条件成立时立即置位并锁存
    IF tankLevel >= 85.0 THEN
        alarmHigh := TRUE;
    ELSIF tempRising THEN
        // 复位沿清除：仅当危险条件已消失才清除
        alarmHigh := FALSE;
    END_IF

    // --- 低液位报警逻辑 ---
    // 危险条件成立时立即置位并锁存
    IF tankLevel <= 15.0 THEN
        alarmLow := TRUE;
    ELSIF tempRising THEN
        // 复位沿清除：仅当危险条件已消失才清除
        alarmLow := FALSE;
    END_IF

    // --- 出口阀控制 ---
    // 低报警锁存期间关闭，其他情况下开启
    outletValveOpen := NOT alarmLow;

    // --- 进料泵控制 ---
    // inletPermit 为 TRUE 且两个报警均为 FALSE 才运行
    IF inletPermit AND NOT alarmHigh AND NOT alarmLow THEN
        pumpRun := TRUE;
    ELSE
        pumpRun := FALSE;
    END_IF

    // 更新上一拍按钮状态
    prevResetBtn := resetBtn;
END_FUNCTION_BLOCK

(* ---- self-easy-02.candidate_02.st ---- *)
FUNCTION_BLOCK FB
VAR_INPUT
    tankLevel    : REAL;      // 储罐液位百分比 0..100
    outletFlow   : REAL;      // 出口流量 m³/h (预留观测接口)
    inletPermit  : BOOL;      // 进料许可
    resetBtn     : BOOL;      // 复位按钮
END_VAR
VAR_OUTPUT
    pumpRun         : BOOL;   // 进料泵运行命令
    alarmHigh       : BOOL;   // 高液位报警
    alarmLow        : BOOL;   // 低液位报警
    outletValveOpen : BOOL;   // 出口阀开命令
END_VAR
VAR
    prevResetBtn : BOOL := FALSE;  // 上拍复位按钮状态
END_VAR

    // 检测复位按钮上升沿：FALSE -> TRUE
    VAR tempRising : BOOL;
    tempRising := resetBtn AND NOT prevResetBtn;

    // --- 高液位报警逻辑 ---
    // 危险条件成立时立即置位并锁存
    IF tankLevel >= 85.0 THEN
        alarmHigh := TRUE;
    ELSIF tempRising THEN
        // 复位沿清除：仅当危险条件已消失才清除
        alarmHigh := FALSE;
    END_IF

    // --- 低液位报警逻辑 ---
    // 危险条件成立时立即置位并锁存
    IF tankLevel <= 15.0 THEN
        alarmLow := TRUE;
    ELSIF tempRising THEN
        // 复位沿清除：仅当危险条件已消失才清除
        alarmLow := FALSE;
    END_IF

    // --- 出口阀控制 ---
    // 低报警锁存期间关闭，其他情况下开启
    outletValveOpen := NOT alarmLow;

    // --- 进料泵控制 ---
    // inletPermit 为 TRUE 且两个报警均为 FALSE 才运行
    IF inletPermit AND NOT alarmHigh AND NOT alarmLow THEN
        pumpRun := TRUE;
    ELSE
        pumpRun := FALSE;
    END_IF

    // 更新上一拍按钮状态
    prevResetBtn := resetBtn;
END_FUNCTION_BLOCK

(* ---- self-hard-01.candidate_01.st ---- *)
FUNCTION_BLOCK FB
VAR_INPUT
    flowLow   : BOOL;
    ackBtn    : BOOL;
    sensorOK  : BOOL;
END_VAR

VAR_OUTPUT
    alarmActive : BOOL;
    alarmAcked  : BOOL;
    highHigh    : BOOL;
END_VAR

VAR
    prev_ackBtn   : BOOL;    (* Previous cycle ackBtn state for rising edge detection *)
END_VAR

VAR_TEMP
    rising_ackBtn : BOOL;    (* Rising edge of ackBtn in current cycle *)
END_VAR

// Detect rising edge of acknowledge button
rising_ackBtn := ackBtn AND NOT prev_ackBtn;

// S5: High priority alarm - sensor failure
highHigh := NOT sensorOK;

// Low priority alarm state machine
// Priority: reset alarmAcked on new flowLow > acknowledge on rising edge > clear on condition gone + acknowledged

IF flowLow THEN
    // Condition occurred: activate alarm, reset acknowledgment
    alarmActive := TRUE;
    alarmAcked := FALSE;

ELSIF rising_ackBtn AND alarmActive THEN
    // Acknowledge button pressed while alarm active
    alarmAcked := TRUE;

ELSIF NOT flowLow AND alarmAcked THEN
    // Condition cleared and already acknowledged: clear alarm
    alarmActive := FALSE;
    alarmAcked := FALSE;

END_IF;

// Update previous state for next cycle
prev_ackBtn := ackBtn;

END_FUNCTION_BLOCK

(* ---- self-hard-01.candidate_02.st ---- *)
FUNCTION_BLOCK FB
VAR_INPUT
    flowLow   : BOOL;
    ackBtn    : BOOL;
    sensorOK  : BOOL;
END_VAR

VAR_OUTPUT
    alarmActive : BOOL;
    alarmAcked  : BOOL;
    highHigh    : BOOL;
END_VAR

VAR
    prev_ackBtn : BOOL;
END_VAR

VAR_TEMP
    rising_ackBtn : BOOL;
END_VAR

rising_ackBtn := ackBtn AND NOT prev_ackBtn;

// S5: High priority alarm - sensor failure
highHigh := NOT sensorOK;

// Low priority alarm state machine
IF flowLow THEN
    // Condition present: activate alarm, reset acknowledgment
    alarmActive := TRUE;
    alarmAcked := FALSE;

ELSIF rising_ackBtn AND alarmActive THEN
    // Acknowledge button pressed while alarm active: mark acknowledged
    alarmAcked := TRUE;

ELSIF alarmActive AND alarmAcked THEN
    // Condition cleared and already acknowledged: clear alarm
    alarmActive := FALSE;
    alarmAcked := FALSE;

END_IF;

prev_ackBtn := ackBtn;

END_FUNCTION_BLOCK

(* ---- self-hard-02.candidate_01.st ---- *)
FUNCTION_BLOCK FB
VAR_INPUT
    startBtn    : BOOL;
    abortBtn    : BOOL;
    setpoint    : REAL;
    pv          : REAL;
    maxDuration : INT;
END_VAR
VAR_OUTPUT
    elapsed  : INT;
    phase    : INT;
    timeout  : BOOL;
END_VAR
VAR
    prev_startBtn : BOOL := FALSE;
    prev_phase    : INT  := 0;
END_VAR

; Save previous values at start of each scan cycle
prev_startBtn := startBtn;
prev_phase    := phase;

; Priority: abort > new start edge > running count
; Highest priority: abortBtn immediately transitions to phase=9
IF abortBtn THEN
    phase := 9;
    ; elapsed and timeout remain unchanged from previous scan

; No abort: check for new start rising edge
ELSIF startBtn AND NOT prev_startBtn THEN
    phase    := 1;
    elapsed  := 0;
    timeout  := FALSE;

; Normal operation: no abort, no new start edge
ELSE
    ; Running phases (1 or 2) accumulate scan counts
    IF prev_phase = 1 OR prev_phase = 2 THEN
        elapsed := elapsed + 1;

        ; Check timeout condition (takes priority over pv-based transition)
        IF elapsed >= maxDuration THEN
            timeout := TRUE;
            phase   := 3;
        ; pv-based phase transition when not timed out
        ELSIF pv >= setpoint THEN
            phase := 2;
        ELSE
            phase := 1;
        END_IF;
    END_IF;

    ; Frozen states (phase=3 or phase=9) keep their values
    ; No action needed - phase, elapsed, timeout retain previous values
END_IF;
END_FUNCTION_BLOCK

(* ---- self-hard-02.candidate_02.st ---- *)
FUNCTION_BLOCK FB
VAR_INPUT
    startBtn    : BOOL;
    abortBtn    : BOOL;
    setpoint    : REAL;
    pv          : REAL;
    maxDuration : INT;
END_VAR
VAR_OUTPUT
    elapsed  : INT;
    phase    : INT;
    timeout  : BOOL;
END_VAR
VAR
    prev_startBtn : BOOL := FALSE;
    prev_phase    : INT  := 0;
END_VAR

prev_startBtn := startBtn;
prev_phase    := phase;

IF abortBtn THEN
    phase := 9;
ELSIF startBtn AND NOT prev_startBtn THEN
    phase   := 1;
    elapsed := 0;
    timeout := FALSE;
ELSE
    IF prev_phase = 1 OR prev_phase = 2 THEN
        elapsed := elapsed + 1;
        IF elapsed >= maxDuration THEN
            timeout := TRUE;
            phase   := 3;
        ELSIF pv >= setpoint THEN
            phase := 2;
        ELSE
            phase := 1;
        END_IF;
    END_IF;
END_IF;
END_FUNCTION_BLOCK

(* ---- self-hard-03.candidate_01.st ---- *)
FUNCTION_BLOCK FB
VAR_INPUT
    pushEn  : BOOL;
    pushItem: INT;
    popEn   : BOOL;
END_VAR

VAR_IN_OUT
    fifo : ARRAY[1..8] OF INT;
END_VAR

VAR_OUTPUT
    count : INT;
    full  : BOOL;
    empty : BOOL;
    head  : INT;
END_VAR

VAR
    prevPushEn : BOOL := FALSE;
    prevPopEn  : BOOL := FALSE;
END_VAR

// ---------------------------------------------------------------------------
// Rising edge detection
// ---------------------------------------------------------------------------
VAR
    risingPush : BOOL;
    risingPop  : BOOL;
END_VAR

risingPush := pushEn AND NOT prevPushEn;
risingPop  := popEn  AND NOT prevPopEn;

// ---------------------------------------------------------------------------
// FIFO logic: pop first, then push
// ---------------------------------------------------------------------------

// 1) Pop on rising edge (non-empty only)
IF risingPop AND count > 0 THEN
    FOR i := 1 TO count - 1 DO
        fifo[i] := fifo[i + 1];
    END_FOR;
    count := count - 1;
END_IF;

// 2) Push on rising edge (only if space available)
IF risingPush AND count < 8 THEN
    count        := count + 1;
    fifo[count]  := pushItem;
END_IF;

// ---------------------------------------------------------------------------
// Outputs
// ---------------------------------------------------------------------------
full  := (count = 8);
empty := (count = 0);

IF count = 0 THEN
    head := 0;
ELSE
    head := fifo[1];
END_IF;

// ---------------------------------------------------------------------------
// Save button histories for next cycle
// ---------------------------------------------------------------------------
prevPushEn := pushEn;
prevPopEn  := popEn;

END_FUNCTION_BLOCK

(* ---- self-hard-03.candidate_02.st ---- *)
FUNCTION_BLOCK FB
VAR_INPUT
    pushEn  : BOOL;
    pushItem: INT;
    popEn   : BOOL;
END_VAR

VAR_IN_OUT
    fifo : ARRAY[1..8] OF INT;
END_VAR

VAR_OUTPUT
    count : INT;
    full  : BOOL;
    empty : BOOL;
    head  : INT;
END_VAR

VAR
    prevPushEn : BOOL := FALSE;
    prevPopEn  : BOOL := FALSE;
    i          : INT;
END_VAR

// ---------------------------------------------------------------------------
// Rising edge detection
// ---------------------------------------------------------------------------
VAR
    risingPush : BOOL;
    risingPop  : BOOL;
END_VAR

risingPush := pushEn AND NOT prevPushEn;
risingPop  := popEn  AND NOT prevPopEn;

// ---------------------------------------------------------------------------
// FIFO logic: pop first, then push
// ---------------------------------------------------------------------------

// 1) Pop on rising edge (non-empty only)
IF risingPop AND count > 0 THEN
    FOR i := 1 TO count - 1 DO
        fifo[i] := fifo[i + 1];
    END_FOR;
    count := count - 1;
END_IF;

// 2) Push on rising edge (only if space available)
IF risingPush AND count < 8 THEN
    count        := count + 1;
    fifo[count]  := pushItem;
END_IF;

// ---------------------------------------------------------------------------
// Outputs
// ---------------------------------------------------------------------------
full  := (count = 8);
empty := (count = 0);

IF count = 0 THEN
    head := 0;
ELSE
    head := fifo[1];
END_IF;

// ---------------------------------------------------------------------------
// Save button histories for next cycle
// ---------------------------------------------------------------------------
prevPushEn := pushEn;
prevPopEn  := popEn;

END_FUNCTION_BLOCK

(* ---- self-hard-04.candidate_01.st ---- *)
FUNCTION_BLOCK FB
VAR_INPUT
    demand     : INT;
    runHours   : ARRAY[1..5] OF LINT;
    rotated    : BOOL;
END_VAR

VAR_OUTPUT
    leadPump   : INT := 0;
    lagPump    : INT := 0;
    runningCount : INT := 0;
END_VAR

VAR
    prevDemand       : INT := 0;
    prevLeadPump     : INT := 0;
    prevLagPump      : INT := 0;
    prevRunningCount : INT := 0;
END_VAR

VAR_TEMP
    clippedDemand : INT;
    minHours      : LINT;
    minPump       : INT;
    minLagHours   : LINT;
    minLagPump    : INT;
    i             : INT;
    hourDiff      : LINT;
END_VAR

// Clip demand to 0..5
clippedDemand := LIMIT(0, demand, 5);
runningCount := clippedDemand;

// Find minimum run hours pump
minHours := runHours[1];
minPump := 1;
FOR i := 2 TO 5 DO
    IF runHours[i] < minHours OR (runHours[i] = minHours AND i < minPump) THEN
        minHours := runHours[i];
        minPump := i;
    END_IF
END_FOR

// Demand = 0: clear pumps
IF clippedDemand = 0 THEN
    leadPump := 0;
    lagPump := 0;
ELSE
    // Demand > 0: select/keep lead pump
    IF prevLeadPump = 0 THEN
        // Initial selection or restart: select minimum (runHours, pumpNumber)
        leadPump := minPump;
    ELSIF rotated AND (runHours[prevLeadPump] - minHours > LINT#50) THEN
        // Hysteresis: only switch if rotated AND gap > 50 hours
        leadPump := minPump;
    ELSE
        // Keep previous lead pump
        leadPump := prevLeadPump;
    END_IF

    // Lag pump selection
    IF clippedDemand >= 2 THEN
        // Need lag pump
        IF lagPump = 0 OR leadPump <> prevLeadPump OR clippedDemand > prevRunningCount THEN
            // Initial selection, main pump changed, or running count increased
            minLagHours := LINT#999999999;
            minLagPump := 0;
            FOR i := 1 TO 5 DO
                IF i <> leadPump THEN
                    IF runHours[i] < minLagHours OR (runHours[i] = minLagHours AND i < minLagPump) THEN
                        minLagHours := runHours[i];
                        minLagPump := i;
                    END_IF
                END_IF
            END_FOR
            lagPump := minLagPump;
        ELSE
            // Keep previous lag pump
            lagPump := prevLagPump;
        END_IF
    ELSE
        lagPump := 0;
    END_IF
END_IF

// Update previous values
prevDemand := clippedDemand;
prevLeadPump := leadPump;
prevLagPump := lagPump;
prevRunningCount := runningCount;

END_FUNCTION_BLOCK

(* ---- self-hard-05.candidate_01.st ---- *)
FUNCTION_BLOCK FB
VAR_INPUT
    runRequest : BOOL;
    flameOK    : BOOL;
    o2Valid    : BOOL;
    o2PV       : REAL;
    baseAir    : REAL;
    resetBtn   : BOOL;
END_VAR

VAR_OUTPUT
    fuelPermit : BOOL;
    trimEnable : BOOL;
    airTrim    : REAL;
    airCommand : REAL;
    tripLatched: BOOL;
    o2Fault    : BOOL;
END_VAR

VAR
    prevResetBtn : BOOL := FALSE;
END_VAR

// ── 熄火跳闸（当拍置位，检测优先于复位）───────────────────────
IF runRequest AND NOT flameOK THEN
    tripLatched := TRUE;
ELSIF resetBtn AND NOT prevResetBtn AND NOT runRequest AND NOT flameOK THEN
    tripLatched := FALSE;
ELSE
    tripLatched := tripLatched;
END_IF

// ── 燃料许可 ───────────────────────────────────────────────────
fuelPermit := runRequest AND flameOK AND NOT tripLatched;

// ── 氧量分析仪故障检测 ─────────────────────────────────────────
o2Fault := NOT o2Valid OR o2PV < 0.0 OR o2PV > 21.0;

// ── 氧量修正投入 ───────────────────────────────────────────────
trimEnable := fuelPermit AND NOT o2Fault;

// ── 氧量修正偏置（钳位 ±10，故障时归零）────────────────────────
IF trimEnable THEN
    airTrim := 2.0 * (2.0 - o2PV);
    IF airTrim > 10.0 THEN
        airTrim := 10.0;
    ELSIF airTrim < -10.0 THEN
        airTrim := -10.0;
    END_IF;
ELSE
    airTrim := 0.0;
END_IF;

// ── 风门命令（燃料许可时叠加修正并钳位 0..100，否则归零）────────
IF fuelPermit THEN
    airCommand := baseAir + airTrim;
    IF airCommand > 100.0 THEN
        airCommand := 100.0;
    ELSIF airCommand < 0.0 THEN
        airCommand := 0.0;
    END_IF;
ELSE
    airCommand := 0.0;
END_IF;

// ── 保存本拍复位按钮状态，供下拍边沿检测 ───────────────────────
prevResetBtn := resetBtn;

END_FUNCTION_BLOCK

(* ---- self-hard-06.candidate_01.st ---- *)
FUNCTION_BLOCK FB
VAR_INPUT
    runRequest      : BOOL;          (* 运行请求 *)
    pressure        : REAL;          (* 母管压力 kPa *)
    pressureValid   : BOOL;          (* 压力变送器数据有效 *)
    fuelFlow        : REAL;          (* 燃料流量 t/h *)
    steamFlow       : REAL;          (* 蒸汽流量 t/h *)
    outletCmd       : INT;           (* 减温减压阀开度命令 % *)
    outletFeedback  : INT;           (* 减温减压阀开度反馈 % *)
    resetBtn        : BOOL;          (* 复位按钮上升沿有效 *)
END_VAR

VAR_OUTPUT
    tripLatched     : BOOL;          (* 超压跳闸自保持 *)
    fuelPermit      : BOOL;          (* 燃料许可 *)
    currentCauseMask: WORD;          (* 本周期诊断线索位掩码 *)
    latchedCauseMask: WORD;          (* 跳闸期间线索累积掩码 *)
    diagnosticActive: BOOL;          (* 存在有效诊断线索 *)
END_VAR

VAR
    prevRunRequest  : BOOL;          (* 上周期 runRequest *)
    prevResetBtn    : BOOL;          (* 上周期 resetBtn *)
    stickyCounter   : INT;           (* 阀卡滞连续周期计数 *)
END_VAR

(* 局部变量 *)
VAR
    risingReset     : BOOL;          (* 复位上升沿 *)
    stickyCondMet   : BOOL;          (* 本拍卡滞输入条件 *)
    stickyCondPrev1 : BOOL;          (* 上一拍卡滞输入条件 *)
    stickyCondPrev2 : BOOL;          (* 上两拍卡滞输入条件 *)
END_VAR

// -------------------------------------------
// 1. 边沿检测
// -------------------------------------------
risingReset := resetBtn AND NOT prevResetBtn;

// -------------------------------------------
// 2. 跳闸条件判断
// -------------------------------------------
IF runRequest AND (NOT pressureValid OR pressure >= 4500.0) THEN
    tripLatched := TRUE;
ELSIF risingReset AND NOT runRequest AND pressureValid AND pressure <= 4200.0 THEN
    tripLatched := FALSE;
END_IF

// -------------------------------------------
// 3. 燃料许可
// -------------------------------------------
fuelPermit := runRequest AND NOT tripLatched;

// -------------------------------------------
// 4. 卡滞连续判据（连续3拍）
// -------------------------------------------
(* 本拍卡滞输入条件：超压工况下阀命令>=50且反馈<=10 *)
stickyCondMet := runRequest AND pressureValid AND (pressure >= 4500.0)
                 AND (outletCmd >= 50) AND (outletFeedback <= 10);

(* 连续性判断：需本拍及此前连续两拍均满足 *)
IF stickyCondMet THEN
    IF stickyCounter < 3 THEN
        stickyCounter := stickyCounter + 1;
    END_IF
ELSE
    stickyCounter := 0;  (* 任一条件不满足立即清零 *)
END_IF

(* 卡滞位成立条件：计数器已达3 *)
VAR
    stickyBitActive : BOOL;
END_VAR
stickyBitActive := (stickyCounter >= 3);

// -------------------------------------------
// 5. 本拍线索掩码计算
// -------------------------------------------
IF NOT runRequest THEN
    (* 无运行请求时线索为0 *)
    currentCauseMask := 0;
ELSIF NOT pressureValid THEN
    (* 变送器失效：bit0=1 *)
    currentCauseMask := 1;
ELSE
    (* 运行中且数据有效 *)
    VAR
        causeVal : INT;
    END_VAR
    causeVal := 0;

    (* bit1: 阀卡滞 *)
    IF stickyBitActive THEN
        causeVal := causeVal + 2;
    END_IF

    (* bit2: 燃烧过剩 *)
    IF (fuelFlow >= 4.0) AND (steamFlow <= 10.0) THEN
        causeVal := causeVal + 4;
    END_IF

    (* 超压但无其他线索：置bit3 *)
    IF (pressure >= 4500.0) AND (causeVal = 0) THEN
        causeVal := 8;
    END_IF

    currentCauseMask := INT_TO_WORD(causeVal);
END_IF

// -------------------------------------------
// 6. 历史线索累积
// -------------------------------------------
IF tripLatched THEN
    latchedCauseMask := latchedCauseMask OR currentCauseMask;
ELSE
    latchedCauseMask := 0;  (* 未跳闸时清零 *)
END_IF

// -------------------------------------------
// 7. 诊断有效位
// -------------------------------------------
diagnosticActive := (currentCauseMask <> 0);

// -------------------------------------------
// 8. 更新状态（供下周期边沿检测和连续性判断）
// -------------------------------------------
prevRunRequest := runRequest;
prevResetBtn   := resetBtn;

END_FUNCTION_BLOCK

(* ---- self-hard-06.candidate_02.st ---- *)
FUNCTION_BLOCK FB
VAR_INPUT
    runRequest      : BOOL;          (* 运行请求 *)
    pressure        : REAL;          (* 母管压力 kPa *)
    pressureValid   : BOOL;          (* 压力变送器数据有效 *)
    fuelFlow        : REAL;          (* 燃料流量 t/h *)
    steamFlow       : REAL;          (* 蒸汽流量 t/h *)
    outletCmd       : INT;           (* 减温减压阀开度命令 % *)
    outletFeedback  : INT;           (* 减温减压阀开度反馈 % *)
    resetBtn        : BOOL;          (* 复位按钮上升沿有效 *)
END_VAR

VAR_OUTPUT
    tripLatched     : BOOL;          (* 超压跳闸自保持 *)
    fuelPermit      : BOOL;          (* 燃料许可 *)
    currentCauseMask: WORD;          (* 本周期诊断线索位掩码 *)
    latchedCauseMask: WORD;          (* 跳闸期间线索累积掩码 *)
    diagnosticActive: BOOL;          (* 存在有效诊断线索 *)
END_VAR

VAR
    prevRunRequest  : BOOL;          (* 上周期 runRequest *)
    prevResetBtn    : BOOL;          (* 上周期 resetBtn *)
    stickyCounter   : INT;           (* 阀卡滞连续周期计数 *)
    risingReset     : BOOL;          (* 复位上升沿 *)
    stickyCondMet   : BOOL;          (* 本拍卡滞输入条件 *)
    causeVal        : INT;           (* 本拍线索计算中间值 *)
END_VAR

// -------------------------------------------
// 1. 边沿检测
// -------------------------------------------
risingReset := resetBtn AND NOT prevResetBtn;

// -------------------------------------------
// 2. 跳闸条件判断
// -------------------------------------------
IF runRequest AND (NOT pressureValid OR pressure >= 4500.0) THEN
    tripLatched := TRUE;
ELSIF risingReset AND NOT runRequest AND pressureValid AND pressure <= 4200.0 THEN
    tripLatched := FALSE;
END_IF

// -------------------------------------------
// 3. 燃料许可
// -------------------------------------------
fuelPermit := runRequest AND NOT tripLatched;

// -------------------------------------------
// 4. 卡滞连续判据（连续3拍）
// -------------------------------------------
(* 本拍卡滞输入条件：超压工况下阀命令>=50且反馈<=10 *)
stickyCondMet := runRequest AND pressureValid AND (pressure >= 4500.0)
                 AND (outletCmd >= 50) AND (outletFeedback <= 10);

(* 连续性判断：需本拍及此前连续两拍均满足 *)
IF stickyCondMet THEN
    IF stickyCounter < 3 THEN
        stickyCounter := stickyCounter + 1;
    END_IF
ELSE
    stickyCounter := 0;  (* 任一条件不满足立即清零 *)
END_IF

// -------------------------------------------
// 5. 本拍线索掩码计算
// -------------------------------------------
IF NOT runRequest THEN
    (* 无运行请求时线索为0 *)
    currentCauseMask := 0;
    causeVal := 0;
ELSIF NOT pressureValid THEN
    (* 变送器失效：bit0=1 *)
    currentCauseMask := 1;
    causeVal := 0;
ELSE
    (* 运行中且数据有效 *)
    causeVal := 0;

    (* bit1: 阀卡滞（连续3拍） *)
    IF stickyCounter >= 3 THEN
        causeVal := causeVal + 2;
    END_IF

    (* bit2: 燃烧过剩 *)
    IF (fuelFlow >= 4.0) AND (steamFlow <= 10.0) THEN
        causeVal := causeVal + 4;
    END_IF

    (* 超压但无其他线索：置bit3 *)
    IF (pressure >= 4500.0) AND (causeVal = 0) THEN
        causeVal := 8;
    END_IF

    currentCauseMask := INT_TO_WORD(causeVal);
END_IF

// -------------------------------------------
// 6. 历史线索累积
// -------------------------------------------
IF tripLatched THEN
    latchedCauseMask := latchedCauseMask OR currentCauseMask;
ELSE
    latchedCauseMask := 0;  (* 未跳闸时清零 *)
END_IF

// -------------------------------------------
// 7. 诊断有效位
// -------------------------------------------
diagnosticActive := (currentCauseMask <> 0);

// -------------------------------------------
// 8. 更新状态（供下周期边沿检测和连续性判断）
// -------------------------------------------
prevRunRequest := runRequest;
prevResetBtn   := resetBtn;

END_FUNCTION_BLOCK

(* ---- self-hard-07.candidate_01.st ---- *)
FUNCTION_BLOCK FB
VAR_INPUT
    mode            : INT;
    resetBtn        : BOOL;
    scanSeconds     : REAL;
    tempSP          : REAL;
    tempPV          : REAL;
    flowPV          : REAL;
    manualFlowSP    : REAL;
    manualValve     : REAL;
END_VAR
VAR_OUTPUT
    flowSP          : REAL;
    valveCommand    : REAL;
    fault           : BOOL;
    normalMode      : BOOL;
END_VAR
VAR
    prevResetBtn    : BOOL := FALSE;
    prevMode        : INT;
    firstScan       : BOOL := TRUE;
    accT            : REAL := 0.0;
    accF            : REAL := 0.0;
    prevValveCommand: REAL := 0.0;
END_VAR

VAR
    eT              : REAL;
    eF              : REAL;
    trial           : REAL;
END_VAR

// Initialize outputs on first scan
IF firstScan THEN
    flowSP := manualFlowSP;
    valveCommand := manualValve;
    firstScan := FALSE;
END_IF

// Fault detection
fault := (mode < 0) OR (mode > 2) OR (scanSeconds <= 0.0) OR (scanSeconds > 10.0);

// Detect rising edge of resetBtn
IF resetBtn AND NOT prevResetBtn THEN
    // Reset action - back to initial state
    flowSP := manualFlowSP;
    valveCommand := manualValve;
    accT := 0.0;
    accF := 0.0;
    normalMode := FALSE;
ELSIF fault THEN
    // Fault fallback - immediate follow manual, no integration, preset integrators
    flowSP := manualFlowSP;
    valveCommand := manualValve;
    accT := 0.0;
    accF := 0.0;
    normalMode := FALSE;
ELSE
    // Mode switch detection (not first scan, no fault, no reset rising edge)
    IF firstScan = FALSE AND mode <> prevMode THEN
        // Bumpless transfer on mode change
        IF mode = 2 THEN
            // Switch to cascade: both outputs keep previous values
            flowSP := flowSP;
            valveCommand := valveCommand;
        ELSE
            // Switch to auto/manual: flowSP follows manual, valve keeps previous
            flowSP := manualFlowSP;
            valveCommand := valveCommand;
        END_IF
        prevMode := mode;
        normalMode := FALSE;
    ELSE
        // Check normal mode condition
        // normalMode = TRUE when: not first scan, mode unchanged, no fault, no reset rising edge
        normalMode := (firstScan = FALSE) AND (mode = prevMode) AND NOT fault AND NOT (resetBtn AND NOT prevResetBtn);

        IF normalMode THEN
            // Normal PI calculation
            // Outer loop: Temperature -> FlowSP
            eT := tempSP - tempPV;
            trial := accT + 0.2 * eT * scanSeconds;
            flowSP := LIMIT(0.0, 1.0 * eT + trial, 50.0);
            accT := flowSP - 1.0 * eT;

            // Inner loop: Flow -> Valve
            eF := flowSP - flowPV;
            trial := accF + 0.5 * eF * scanSeconds;
            valveCommand := LIMIT(0.0, 2.0 * eF + trial, 100.0);
            accF := valveCommand - 2.0 * eF;
        END_IF
    END_IF
END_IF

// Update previous cycle variables
prevMode := mode;
prevResetBtn := resetBtn;
prevValveCommand := valveCommand;
END_FUNCTION_BLOCK

(* ---- self-hard-07.candidate_02.st ---- *)
FUNCTION_BLOCK FB
VAR_INPUT
    mode            : INT;
    resetBtn        : BOOL;
    scanSeconds     : REAL;
    tempSP          : REAL;
    tempPV          : REAL;
    flowPV          : REAL;
    manualFlowSP    : REAL;
    manualValve     : REAL;
END_VAR
VAR_OUTPUT
    flowSP          : REAL;
    valveCommand    : REAL;
    fault           : BOOL;
    normalMode      : BOOL;
END_VAR
VAR
    prevResetBtn        : BOOL := FALSE;
    prevMode            : INT := 999;
    firstCycle          : BOOL := TRUE;
    initialized         : BOOL := FALSE;
    accT                : REAL := 0.0;
    accF                : REAL := 0.0;
    prevTempSP          : REAL := 0.0;
    prevTempPV          : REAL := 0.0;
    prevFlowSP          : REAL := 0.0;
    prevValveCommand    : REAL := 0.0;
END_VAR

VAR
    eT      : REAL;
    eF      : REAL;
    trial   : REAL;
END_VAR

eT := tempSP - tempPV;
eF := flowSP - flowPV;

IF firstCycle THEN
    flowSP := manualFlowSP;
    valveCommand := manualValve;
    firstCycle := FALSE;
    initialized := TRUE;
    normalMode := FALSE;
    prevMode := mode;
    prevResetBtn := resetBtn;
    prevTempSP := tempSP;
    prevTempPV := tempPV;
    prevFlowSP := flowSP;
    prevValveCommand := valveCommand;
    RETURN;
END_IF;

fault := (mode < 0) OR (mode > 2) OR (scanSeconds <= 0.0) OR (scanSeconds > 10.0);

IF resetBtn AND NOT prevResetBtn THEN
    flowSP := manualFlowSP;
    valveCommand := manualValve;
    accT := 0.0;
    accF := 0.0;
    normalMode := FALSE;
    prevMode := mode;
    prevResetBtn := resetBtn;
    prevTempSP := tempSP;
    prevTempPV := tempPV;
    prevFlowSP := flowSP;
    prevValveCommand := valveCommand;
    RETURN;
END_IF;

IF fault THEN
    flowSP := manualFlowSP;
    valveCommand := manualValve;
    accT := 0.0;
    accF := 0.0;
    normalMode := FALSE;
    prevMode := mode;
    prevResetBtn := resetBtn;
    prevTempSP := tempSP;
    prevTempPV := tempPV;
    prevFlowSP := flowSP;
    prevValveCommand := valveCommand;
    RETURN;
END_IF;

IF mode <> prevMode THEN
    IF mode = 2 THEN
        flowSP := prevFlowSP;
        valveCommand := prevValveCommand;
    ELSE
        flowSP := manualFlowSP;
    END_IF;
    normalMode := FALSE;
    prevMode := mode;
    prevResetBtn := resetBtn;
    prevTempSP := tempSP;
    prevTempPV := tempPV;
    prevFlowSP := flowSP;
    prevValveCommand := valveCommand;
    RETURN;
END_IF;

normalMode := TRUE;

trial := accT + 0.2 * eT * scanSeconds;
flowSP := LIMIT(0.0, 1.0 * eT + trial, 50.0);
accT := flowSP - 1.0 * eT;

trial := accF + 0.5 * eF * scanSeconds;
valveCommand := LIMIT(0.0, 2.0 * eF + trial, 100.0);
accF := valveCommand - 2.0 * eF;

prevTempSP := tempSP;
prevTempPV := tempPV;
prevFlowSP := flowSP;
prevValveCommand := valveCommand;
prevResetBtn := resetBtn;
prevMode := mode;
END_FUNCTION_BLOCK

(* ---- self-medium-01.candidate_01.st ---- *)
FUNCTION_BLOCK FB
VAR_INPUT
    recipe: ARRAY[1..8] OF ST_Recipe;
    selSlot: INT;
    loadCmd: BOOL;
    running: BOOL;
END_VAR

VAR_OUTPUT
    valid: BOOL;
    loadedID: INT;
END_VAR

VAR
    prevLoadCmd: BOOL := FALSE;
    prevLoadedID: INT := 0;
    prevValid: BOOL := FALSE;
END_VAR

VAR
    risingEdge: BOOL;
END_VAR

risingEdge := loadCmd AND NOT prevLoadCmd;

IF risingEdge AND NOT running THEN
    IF (selSlot >= 1) AND (selSlot <= 8) THEN
        IF (recipe[selSlot].recipeID <> 0) AND
           (recipe[selSlot].totalRatio >= 99.0) AND
           (recipe[selSlot].totalRatio <= 101.0) AND
           (recipe[selSlot].temperature >= 30.0) AND
           (recipe[selSlot].temperature <= 180.0) THEN
            loadedID := recipe[selSlot].recipeID;
            valid := TRUE;
        ELSE
            loadedID := 0;
            valid := FALSE;
        END_IF
    ELSE
        loadedID := 0;
        valid := FALSE;
    END_IF;
ELSE
    loadedID := prevLoadedID;
    valid := prevValid;
END_IF;

prevLoadedID := loadedID;
prevValid := valid;
prevLoadCmd := loadCmd;

(* ---- self-medium-01.candidate_02.st ---- *)
TYPE ST_Recipe :
STRUCT
    recipeID: INT;
    totalRatio: REAL;
    temperature: REAL;
END_STRUCT
END_TYPE

FUNCTION_BLOCK FB
VAR_INPUT
    recipe: ARRAY[1..8] OF ST_Recipe;
    selSlot: INT;
    loadCmd: BOOL;
    running: BOOL;
END_VAR

VAR_OUTPUT
    valid: BOOL;
    loadedID: INT;
END_VAR

VAR
    prevLoadCmd: BOOL := FALSE;
    prevLoadedID: INT := 0;
    prevValid: BOOL := FALSE;
    risingEdge: BOOL;
END_VAR

risingEdge := loadCmd AND NOT prevLoadCmd;

IF risingEdge AND NOT running THEN
    IF (selSlot >= 1) AND (selSlot <= 8) THEN
        IF (recipe[selSlot].recipeID <> 0) AND
           (recipe[selSlot].totalRatio >= 99.0) AND
           (recipe[selSlot].totalRatio <= 101.0) AND
           (recipe[selSlot].temperature >= 30.0) AND
           (recipe[selSlot].temperature <= 180.0) THEN
            loadedID := recipe[selSlot].recipeID;
            valid := TRUE;
        ELSE
            loadedID := 0;
            valid := FALSE;
        END_IF
    ELSE
        loadedID := 0;
        valid := FALSE;
    END_IF;
ELSE
    IF running THEN
        loadedID := prevLoadedID;
        valid := prevValid;
    END_IF;
END_IF;

prevLoadedID := loadedID;
prevValid := valid;
prevLoadCmd := loadCmd;

END_FUNCTION_BLOCK

(* ---- self-medium-02.candidate_01.st ---- *)
FUNCTION_BLOCK FB
VAR_INPUT
    enable      : BOOL;
    rawValue    : REAL;
END_VAR

VAR_OUTPUT
    filteredValue : REAL := 0.0;
    windowFull    : BOOL := FALSE;
    sampleCount   : INT  := 0;
END_VAR

VAR
    buffer     : ARRAY[0..7] OF REAL;
    writeIndex : INT := 0;
    sum        : REAL;
    i          : INT;
    prev_enable : BOOL := FALSE;
END_VAR

// Initialization on rising edge or first power-up with enable already TRUE
IF enable AND sampleCount = 0 THEN
    writeIndex  := 0;
    sampleCount := 0;
    windowFull  := FALSE;
END_IF;

// Detect rising edge on enable
IF enable AND NOT prev_enable THEN
    writeIndex  := 0;
    sampleCount := 0;
    windowFull  := FALSE;
END_IF;

IF enable THEN
    // Write new sample into circular buffer
    buffer[writeIndex] := rawValue;
    writeIndex := (writeIndex + 1) MOD 8;

    // Increment sample count (cap at 8)
    IF sampleCount < 8 THEN
        sampleCount := sampleCount + 1;
    END_IF;

    // Set windowFull flag when 8 samples accumulated
    IF sampleCount = 8 THEN
        windowFull := TRUE;
    END_IF;

    // Calculate sum of valid samples in circular buffer
    sum := 0.0;
    IF sampleCount = 8 THEN
        // Buffer full: sum all 8 samples (oldest at writeIndex)
        FOR i := 0 TO 7 DO
            sum := sum + buffer[i];
        END_FOR;
        filteredValue := sum / 8.0;
    ELSE
        // Buffer not full: sum first sampleCount samples
        FOR i := 0 TO sampleCount - 1 DO
            sum := sum + buffer[i];
        END_FOR;
        filteredValue := sum / INT_TO_REAL(sampleCount);
    END_IF;
ELSE
    // enable = FALSE: clear count and full flag, keep filteredValue unchanged
    sampleCount := 0;
    windowFull  := FALSE;
END_IF;

// Track previous enable state for edge detection
prev_enable := enable;
END_FUNCTION_BLOCK

(* ---- self-medium-03.candidate_01.st ---- *)
FUNCTION_BLOCK FB
VAR_INPUT
    openBtn    : BOOL;
    closeBtn   : BOOL;
    openLimit  : BOOL;
    closeLimit : BOOL;
    obstacle   : BOOL;
END_VAR
VAR_OUTPUT
    motorUp    : BOOL;
    motorDown  : BOOL;
    errorFlag  : BOOL;
END_VAR
VAR
    prev_openBtn  : BOOL := FALSE;
    prev_closeBtn : BOOL := FALSE;
    prev_obstacle : BOOL := FALSE;
    // Internal state: 0=IDLE, 1=OPENING, 2=CLOSING, 3=FAULT
    state : INT := 0;
END_VAR
VAR
    risingEdgeOpen  : BOOL;
    risingEdgeClose : BOOL;
    risingEdgeBoth  : BOOL;
END_VAR

// ============================================================================
// Edge Detection
// ============================================================================
risingEdgeOpen  := openBtn  AND NOT prev_openBtn;
risingEdgeClose := closeBtn AND NOT prev_closeBtn;
risingEdgeBoth  := (openBtn AND closeBtn) AND NOT (prev_openBtn AND prev_closeBtn);

// ============================================================================
// Fault Handling (highest priority)
// ============================================================================
IF obstacle THEN
    errorFlag := TRUE;
    state := 3; // FAULT
END_IF;

// ============================================================================
// State Transitions & Motor Control
// ============================================================================
CASE state OF
    // ---- IDLE ----
    0: // IDLE
        IF errorFlag THEN
            // Already in fault, stay here
            motorUp   := FALSE;
            motorDown := FALSE;
        ELSE
            // Check for new open command
            IF risingEdgeOpen AND NOT closeBtn AND NOT openLimit AND NOT obstacle THEN
                state     := 1; // OPENING
                motorUp   := TRUE;
                motorDown := FALSE;
            // Check for new close command
            ELSIF risingEdgeClose AND NOT openBtn AND NOT closeLimit AND NOT obstacle THEN
                state     := 2; // CLOSING
                motorUp   := FALSE;
                motorDown := TRUE;
            ELSE
                motorUp   := FALSE;
                motorDown := FALSE;
            END_IF;
        END_IF;

    // ---- OPENING ----
    1: // OPENING
        IF obstacle THEN
            // Handled above, stay in fault
            motorUp   := FALSE;
            motorDown := FALSE;
        ELSIF openLimit THEN
            state     := 0; // IDLE
            motorUp   := FALSE;
            motorDown := FALSE;
        ELSE
            // Continue opening
            motorUp   := TRUE;
            motorDown := FALSE;
        END_IF;

    // ---- CLOSING ----
    2: // CLOSING
        IF obstacle THEN
            // Handled above, stay in fault
            motorUp   := FALSE;
            motorDown := FALSE;
        ELSIF closeLimit THEN
            state     := 0; // IDLE
            motorUp   := FALSE;
            motorDown := FALSE;
        ELSE
            // Continue closing
            motorUp   := FALSE;
            motorDown := TRUE;
        END_IF;

    // ---- FAULT ----
    3: // FAULT
        motorUp   := FALSE;
        motorDown := FALSE;
        // Reset only when no obstacle AND both buttons have new rising edge together
        IF NOT obstacle AND risingEdgeBoth THEN
            errorFlag := FALSE;
            state     := 0; // IDLE
        END_IF;
END_CASE;

// ============================================================================
// Update Previous States for Next Scan
// ============================================================================
prev_openBtn  := openBtn;
prev_closeBtn := closeBtn;
prev_obstacle := obstacle;

END_FUNCTION_BLOCK

(* ---- self-medium-04.candidate_01.st ---- *)
FUNCTION_BLOCK FB
VAR_INPUT
    startBtn   : BOOL;
    resetBtn   : BOOL;
    doneSensor : BOOL;
    targetVol  : REAL;
    flowVol    : REAL;
END_VAR
VAR_OUTPUT
    valveOpen  : BOOL;
    fillsToday : INT := 0;
END_VAR
VAR
    prevStartBtn   : BOOL := FALSE;
    prevResetBtn   : BOOL := FALSE;
    prevValveOpen  : BOOL := FALSE;
    prevDoneSensor : BOOL := FALSE;
    prevFillsToday : INT  := 0;

    currentVolume  : REAL := 0.0;
    pendingConfirm : BOOL := FALSE;
END_VAR

VAR_TEMP
    risingStart  : BOOL;
    risingReset  : BOOL;
    risingDone   : BOOL;
END_VAR

// 检测上升沿
risingStart  := startBtn AND NOT prevStartBtn;
risingReset  := resetBtn AND NOT prevResetBtn;
risingDone   := doneSensor AND NOT prevDoneSensor;

// ========== 1. 复位优先 ==========
IF risingReset THEN
    // 清零计数和累计体积
    fillsToday      := 0;
    currentVolume   := 0.0;
    // 关阀并清除待确认
    valveOpen       := FALSE;
    pendingConfirm  := FALSE;
ELSE
    // ========== 2. 启动新瓶 ==========
    IF risingStart THEN
        // 若上一瓶仍待确认，先取消
        pendingConfirm := FALSE;
        // 清零本瓶累计并开阀
        currentVolume  := 0.0;
        valveOpen      := TRUE;
    END_IF;

    // ========== 3. 灌装累计与关阀 ==========
    IF valveOpen THEN
        // 加入本拍流量，启动拍也计入
        currentVolume := currentVolume + flowVol;

        // 累计达到或超过目标时立即关阀并令本瓶待确认
        IF currentVolume >= targetVol THEN
            valveOpen      := FALSE;
            pendingConfirm := TRUE;
        END_IF;
    END_IF;

    // ========== 4. 确认逻辑 ==========
    IF pendingConfirm THEN
        // 本拍关阀后立即读取 doneSensor
        IF doneSensor THEN
            // 本拍确认并计数
            pendingConfirm := FALSE;

            // fillsToday 增加 1；原计数为 32767 时保持 32767
            IF fillsToday < 32767 THEN
                fillsToday := fillsToday + 1;
            END_IF;
        END_IF;
    END_IF;
END_IF;

// 更新上电前值（用于下一拍上升沿检测）
prevStartBtn   := startBtn;
prevResetBtn   := resetBtn;
prevValveOpen  := valveOpen;
prevDoneSensor := doneSensor;
prevFillsToday := fillsToday;
END_FUNCTION_BLOCK

(* ---- self-medium-04.candidate_02.st ---- *)
FUNCTION_BLOCK FB
VAR_INPUT
    startBtn   : BOOL;
    resetBtn   : BOOL;
    doneSensor : BOOL;
    targetVol  : REAL;
    flowVol    : REAL;
END_VAR
VAR_OUTPUT
    valveOpen  : BOOL;
    fillsToday : INT := 0;
END_VAR
VAR
    prevStartBtn   : BOOL := FALSE;
    prevResetBtn   : BOOL := FALSE;
    prevValveOpen  : BOOL := FALSE;

    currentVolume  : REAL := 0.0;
    pendingConfirm : BOOL := FALSE;
END_VAR

VAR_TEMP
    risingStart : BOOL;
    risingReset : BOOL;
END_VAR

risingStart := startBtn AND NOT prevStartBtn;
risingReset := resetBtn AND NOT prevResetBtn;

// ========== 1. 复位优先 ==========
IF risingReset THEN
    fillsToday      := 0;
    currentVolume   := 0.0;
    valveOpen       := FALSE;
    pendingConfirm  := FALSE;
    prevStartBtn    := resetBtn;
    prevResetBtn    := resetBtn;
    RETURN;
END_IF;

// ========== 2. 启动新瓶 ==========
IF risingStart THEN
    pendingConfirm := FALSE;
    currentVolume  := 0.0;

    IF flowVol >= targetVol THEN
        // 启动拍直接达标：关阀，本拍确认
        valveOpen      := FALSE;
        pendingConfirm := TRUE;
    ELSE
        valveOpen := TRUE;
    END_IF;
ELSE
    // ========== 3. 灌装累计 ==========
    IF valveOpen THEN
        currentVolume := currentVolume + flowVol;

        IF currentVolume >= targetVol THEN
            valveOpen      := FALSE;
            pendingConfirm := TRUE;
        END_IF;
    END_IF;
END_IF;

// ========== 4. 确认逻辑 ==========
IF pendingConfirm AND doneSensor THEN
    pendingConfirm := FALSE;
    IF fillsToday < 32767 THEN
        fillsToday := fillsToday + 1;
    END_IF;
END_IF;

prevStartBtn  := startBtn;
prevResetBtn  := resetBtn;
prevValveOpen := valveOpen;
END_FUNCTION_BLOCK

(* ---- self-medium-05.candidate_01.st ---- *)
FUNCTION_BLOCK FB
VAR_INPUT
    enable       : BOOL;
    resetBtn     : BOOL;
    scanSeconds  : LREAL;  // renamed from dt, unit: s
    steamFlow    : LREAL;  // kg/s, valid range [0, 90]
    fuelFlow     : LREAL;  // kg/s, valid range [0, 6]
    steamTemp    : LREAL;  // °C, qualified [447, 453]
    steamPressure: LREAL;  // kPa, qualified [3750, 3850]
END_VAR

VAR_OUTPUT
    qualified    : BOOL;
    dataFault    : BOOL;
    qualifiedTon : LREAL;
    fuelTon      : LREAL;
    revenue      : LREAL;
    cost         : LREAL;
    netProfit    : LREAL;
END_VAR

VAR
    prevResetBtn : BOOL := FALSE;
END_VAR

// Detect rising edge of resetBtn (edge-triggered, not level-triggered)
VAR_TEMP
    risingReset : BOOL;
END_VAR

risingReset := resetBtn AND NOT prevResetBtn;

// Data fault: invalid scan time or out-of-range flow values
dataFault := (scanSeconds <= 0.0 OR scanSeconds > 10.0 OR
              steamFlow < 0.0 OR steamFlow > 90.0 OR
              fuelFlow < 0.0 OR fuelFlow > 6.0);

// Qualified: closed interval [447, 453] °C and [3750, 3850] kPa
qualified := (steamTemp >= 447.0 AND steamTemp <= 453.0) AND
             (steamPressure >= 3750.0 AND steamPressure <= 3850.0);

// Accumulation with priority: reset > enable/fault-free
IF risingReset THEN
    // Reset takes priority; fault flag still reports but accumulators clear
    qualifiedTon := 0.0;
    fuelTon := 0.0;
ELSIF enable AND NOT dataFault THEN
    // Fuel: always accumulate when enabled and data valid
    fuelTon := fuelTon + fuelFlow * scanSeconds / 1000.0;
    // Qualified steam: only when qualified
    IF qualified THEN
        qualifiedTon := qualifiedTon + steamFlow * scanSeconds / 1000.0;
    END_IF;
END_IF;
// When disabled or faulted (without reset), accumulators hold previous values

// Financial calculations (update every scan regardless of accumulation)
revenue   := qualifiedTon * 280.0;  // yuan/t steam
cost      := fuelTon * 1500.0;      // yuan/t fuel
netProfit := revenue - cost;        // may be negative

// Update edge-detection state for next cycle
prevResetBtn := resetBtn;

END_FUNCTION_BLOCK

(* ---- self-medium-06.candidate_01.st ---- *)
FUNCTION_BLOCK FB
VAR_INPUT
    enable         : BOOL;
    resetBtn       : BOOL;
    sensorValid    : BOOL;
    setpoint       : REAL;
    temperature    : REAL;
    scanSeconds    : REAL;
    bias           : REAL;
END_VAR

VAR_OUTPUT
    power      : REAL;
    correction : REAL;
    fault      : BOOL;
END_VAR

VAR
    ePrev       : REAL := 0.0;
    hasHistory  : BOOL := FALSE;
    prevResetBtn : BOOL := FALSE;
END_VAR

// Temp vars
VAR
    e, de, x, y         : REAL;
    muNx, muZx, muPx    : REAL;
    muNy, muZy, muPy    : REAL;
    w_NN, w_NZ, w_NP    : REAL;
    w_ZN, w_ZZ, w_ZP    : REAL;
    w_PN, w_PZ, w_PP    : REAL;
    sumWc, sumW         : REAL;
    resetRising         : BOOL;
END_VAR

// Fault detection
fault := (NOT sensorValid) OR (scanSeconds <= 0.0) OR (scanSeconds > 10.0);

// Rising edge of resetBtn
resetRising := resetBtn AND (NOT prevResetBtn);
prevResetBtn := resetBtn;

// Clear outputs and history on disable, fault, or reset rising edge
IF (NOT enable) OR fault OR resetRising THEN
    power      := 0.0;
    correction := 0.0;
    ePrev      := 0.0;
    hasHistory := FALSE;
ELSE
    // Calculate error
    e := setpoint - temperature;

    // Calculate derivative of error
    // First scan after history cleared: de = 0
    IF hasHistory THEN
        de := (e - ePrev) / scanSeconds;
    ELSE
        de := 0.0;
    END_IF;

    // Normalize error and derivative
    // x range: [-1, 1] for e in [-10, 10] degC
    // y range: [-1, 1] for de in [-2, 2] degC/s
    x := e / 10.0;
    IF x > 1.0 THEN x := 1.0; END_IF;
    IF x < -1.0 THEN x := -1.0; END_IF;

    y := de / 2.0;
    IF y > 1.0 THEN y := 1.0; END_IF;
    IF y < -1.0 THEN y := -1.0; END_IF;

    // Membership functions for x (error)
    muNx := -x;
    IF muNx < 0.0 THEN muNx := 0.0; END_IF;
    muZx := 1.0 - ABS(x);
    muPx := x;
    IF muPx < 0.0 THEN muPx := 0.0; END_IF;

    // Membership functions for y (derivative)
    muNy := -y;
    IF muNy < 0.0 THEN muNy := 0.0; END_IF;
    muZy := 1.0 - ABS(y);
    muPy := y;
    IF muPy < 0.0 THEN muPy := 0.0; END_IF;

    // Rule weights: w(i,j) = mu_i(x) * mu_j(y)
    w_NN := muNx * muNy;  // N x N
    w_NZ := muNx * muZy;  // N x Z
    w_NP := muNx * muPy;  // N x P
    w_ZN := muZx * muNy;  // Z x N
    w_ZZ := muZx * muZy;  // Z x Z
    w_ZP := muZx * muPy;  // Z x P
    w_PN := muPx * muNy;  // P x N
    w_PZ := muPx * muZy;  // P x Z
    w_PP := muPx * muPy;  // P x P

    // Centroid defuzzification
    // Single-point outputs: NxN=-30, NxZ=-20, NxP=-10,
    //                       ZxN=-10, ZxZ=0,   ZxP=10,
    //                       PxN=10,  PxZ=20,  PxP=30
    sumWc := w_NN * (-30.0) + w_NZ * (-20.0) + w_NP * (-10.0)
           + w_ZN * (-10.0) + w_ZZ * 0.0     + w_ZP * 10.0
           + w_PN * 10.0     + w_PZ * 20.0    + w_PP * 30.0;
    sumW := w_NN + w_NZ + w_NP + w_ZN + w_ZZ + w_ZP + w_PN + w_PZ + w_PP;

    IF sumW > 0.0 THEN
        correction := sumWc / sumW;
    ELSE
        correction := 0.0;
    END_IF;

    // Power: bias + correction, clamped to [0, 100]
    power := bias + correction;
    IF power > 100.0 THEN power := 100.0; END_IF;
    IF power < 0.0 THEN power := 0.0; END_IF;

    // Update history for next scan
    ePrev := e;
    hasHistory := TRUE;
END_IF

END_FUNCTION_BLOCK

(* ---- public-easy-01.candidate_01.st ---- *)
PROGRAM FillingLineControl
VAR
    State : INT := 0;  // 0=Idle, 1=Cleaning, 2=Filling, 3=Capping, 4=Packing, 5=Complete
END_VAR

CASE State OF
    0:  // Idle - waiting for bottle
        Pump_Motor := FALSE;
        Filling_Valve := FALSE;
        Capping_Machine := FALSE;
        Packing_Machine := FALSE;
        Completion_Light := FALSE;

        IF bottleSensor THEN
            State := 1;
        END_IF

    1:  // Cleaning
        Pump_Motor := TRUE;

        IF cleaningConfirmButton THEN
            State := 2;
        END_IF

    2:  // Filling
        Pump_Motor := FALSE;
        Filling_Valve := TRUE;

        IF fillingConfirmButton THEN
            State := 3;
        END_IF

    3:  // Capping
        Filling_Valve := FALSE;
        Capping_Machine := TRUE;

        IF cappingConfirmButton THEN
            State := 4;
        END_IF

    4:  // Packing
        Capping_Machine := FALSE;
        Packing_Machine := TRUE;

        IF packingConfirmButton THEN
            State := 5;
        END_IF

    5:  // Complete - packaging finished, waiting for pickup
        Packing_Machine := FALSE;
        Completion_Light := TRUE;

        IF finishedButton THEN
            State := 0;
        END_IF
END_CASE

(* ---- public-easy-01.candidate_02.st ---- *)
PROGRAM FillingLineControl
VAR
    State : INT := 0;  // 0=Idle, 1=Cleaning, 2=Filling, 3=Capping, 4=Packing, 5=Complete
END_VAR

CASE State OF
    0:  // Idle - waiting for bottle
        Pump_Motor := FALSE;
        Filling_Valve := FALSE;
        Capping_Machine := FALSE;
        Packing_Machine := FALSE;
        Completion_Light := FALSE;

        IF bottleSensor THEN
            State := 1;
        END_IF

    1:  // Cleaning
        Pump_Motor := TRUE;

        IF cleaningConfirmButton THEN
            State := 2;
        END_IF

    2:  // Filling
        Pump_Motor := FALSE;
        Filling_Valve := TRUE;

        IF fillingConfirmButton THEN
            State := 3;
        END_IF

    3:  // Capping
        Filling_Valve := FALSE;
        Capping_Machine := TRUE;

        IF cappingConfirmButton THEN
            State := 4;
        END_IF

    4:  // Packing
        Capping_Machine := FALSE;
        Packing_Machine := TRUE;

        IF packingConfirmButton THEN
            State := 5;
        END_IF

    5:  // Complete - packaging finished, waiting for pickup
        Packing_Machine := FALSE;
        Completion_Light := TRUE;

        IF finishedButton THEN
            State := 0;
        END_IF
END_CASE

END_PROGRAM

(* ---- public-easy-04.candidate_01.st ---- *)
PROGRAM JamPumpControl
VAR
    ViscosityDebounceTimer : TON;
    ViscosityConditionValid : BOOL := FALSE;
END_VAR

// Power-up initialization
IF __SYSTEM__:*FIRSTSCAN THEN
    VFD_RUN := FALSE;
    PUMP_RUNTIME_ACC := LTIME#0s;
    PUMP_MAINT_DUE := FALSE;
    ViscosityConditionValid := FALSE;
END_IF;

// Viscosity debouncing logic
// Invalidate immediately when input becomes FALSE
IF NOT VISCOSITY_OK THEN
    ViscosityConditionValid := FALSE;
    ViscosityDebounceTimer(IN := FALSE);
ELSE
    // Start or continue timing when viscosity is good
    ViscosityDebounceTimer(IN := TRUE, PT := DebounceTime);

    // Condition is valid only after timer completes
    IF ViscosityDebounceTimer.Q THEN
        ViscosityConditionValid := TRUE;
    END_IF;
END_IF;

// Emergency stop and run permission logic
// VFD_RUN allowed only when E-STOP is OK AND viscosity is valid
IF PASTE_E_STOP_NC AND ViscosityConditionValid THEN
    VFD_RUN := TRUE;
ELSE
    VFD_RUN := FALSE;
END_IF;

// Runtime accumulation (accumulates only while VFD_RUN is TRUE)
IF VFD_RUN THEN
    PUMP_RUNTIME_ACC := PUMP_RUNTIME_ACC + CycleTime;
END_IF;

// Maintenance due indication (500 hours)
PUMP_MAINT_DUE := (PUMP_RUNTIME_ACC >= LTIME#500h);

END_PROGRAM
